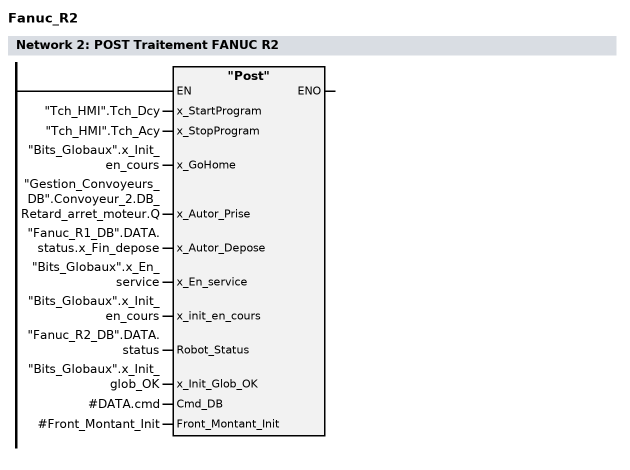
   RUNG wire#powerrail
      "Post"(x_StartProgram := "Tch_HMI".Tch_Dcy, x_StopProgram := "Tch_HMI".Tch_Acy, x_GoHome := "Bits_Globaux".x_Init_en_cours, x_Autor_Prise := "Gestion_Convoyeurs_DB".Convoyeur_2.DB_Retard_arret_moteur.Q, x_Autor_Depose := "Fanuc_R1_DB".DATA.status.x_Fin_depose, x_En_service := "Bits_Globaux".x_En_service, x_init_en_cours := "Bits_Globaux".x_Init_en_cours, Robot_Status := "Fanuc_R2_DB".DATA.status, x_Init_Glob_OK := "Bits_Globaux".x_Init_glob_OK, Cmd_DB := #DATA.cmd, Front_Montant_Init := #Front_Montant_Init)
   END_RUNG
   // the same network as SCL:
   "Post"(x_StartProgram := "Tch_HMI".Tch_Dcy,
          x_StopProgram := "Tch_HMI".Tch_Acy,
          x_GoHome := "Bits_Globaux".x_Init_en_cours,
          x_Autor_Prise := "Gestion_Convoyeurs_DB".Convoyeur_2.DB_Retard_arret_moteur.Q,
          x_Autor_Depose := "Fanuc_R1_DB".DATA.status.x_Fin_depose,
          x_En_service := "Bits_Globaux".x_En_service,
          x_init_en_cours := "Bits_Globaux".x_Init_en_cours,
          Robot_Status := "Fanuc_R2_DB".DATA.status,
          x_Init_Glob_OK := "Bits_Globaux".x_Init_glob_OK,
          Cmd_DB := #DATA.cmd,
          Front_Montant_Init := #Front_Montant_Init);
END_REGION
END_FUNCTION_BLOCK

// folder: 5-Cellule_conditionnement/GoFa_ABB_R3

FUNCTION_BLOCK "GoFa_R3_FB"   // FB15, LAD
TITLE = Commande ABB
{ S7_Optimized_Access := 'TRUE' }
VERSION : 0.1
   VAR
      GoFa_Status : "GoFa_Status";
      GoFa_Cmd : "GoFa_cmd";
      x_Demande_ecriture_Modbus : Bool;
   END_VAR
BEGIN

REGION Network 1: Allumage des moteurs
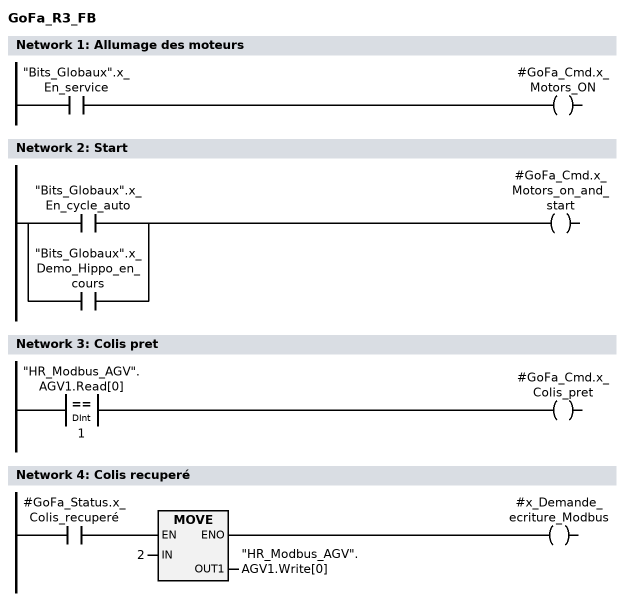
   RUNG wire#powerrail
      Contact( "Bits_Globaux".x_En_service )
      Coil( #GoFa_Cmd.x_Motors_ON )
   END_RUNG
   // the same network as SCL:
   #GoFa_Cmd.x_Motors_ON := "Bits_Globaux".x_En_service;
END_REGION

REGION Network 2: Start
   RUNG wire#powerrail
      Contact( "Bits_Globaux".x_En_cycle_auto )
      wire#w1
      Coil( #GoFa_Cmd.x_Motors_on_and_start )
   END_RUNG
   RUNG wire#powerrail
      Contact( "Bits_Globaux".x_Demo_Hippo_en_cours )
   END_RUNG wire#w1
   // the same network as SCL:
   #GoFa_Cmd.x_Motors_on_and_start := "Bits_Globaux".x_En_cycle_auto OR "Bits_Globaux".x_Demo_Hippo_en_cours;
END_REGION

REGION Network 3: Colis pret
   RUNG wire#powerrail
      { S7_Templates := "SrcType := DInt" } EQ_Contact(in1 := "HR_Modbus_AGV".AGV1.Read[0], in2 := 1)
      Coil( #GoFa_Cmd.x_Colis_pret )
   END_RUNG
   // the same network as SCL:
   #GoFa_Cmd.x_Colis_pret := "HR_Modbus_AGV".AGV1.Read[0] = 1;
END_REGION

REGION Network 4: Colis recuperé
   RUNG wire#powerrail
      Contact( #GoFa_Status.x_Colis_recuperé )
      Move(in := 2, out1 => "HR_Modbus_AGV".AGV1.Write[0])
      Coil( #x_Demande_ecriture_Modbus )
   END_RUNG
   // the same network as SCL:
   IF #GoFa_Status.x_Colis_recuperé THEN "HR_Modbus_AGV".AGV1.Write[0] := 2; END_IF;
   #x_Demande_ecriture_Modbus := #GoFa_Status.x_Colis_recuperé;
END_REGION
END_FUNCTION_BLOCK

// folder: 6_UR10_R5

FUNCTION_BLOCK "60_UR_R5"   // FB6, LAD
{ S7_Optimized_Access := 'TRUE' }
VERSION : 0.1
   VAR
      DATA : "UR_Cobot";
      x_DemandeEcriture_Modbus_AGV : Bool;
   END_VAR
   // // DATA.Registers_Out_2.Bits.Register[0] : Demande Init
   // // DATA.Registers_Out_2.Bits.Register[1] : EnCycleAuto
   // // DATA.Registers_Out_2.Bits.Register[2] : EnCycleDemo
   // // DATA.Registers_Out_2.Bits.Register[3] : PauseProgPLC
   // // DATA.Registers_Out_2.Bits.Register[4] : StopProgPLC
   // // DATA.Registers_Out_2.Bits.Register[5] : StartProgPLC (demarrage boucle Main)
   // // DATA.Registers_Out_2.Bits.Register[6] : Initialisation auto après AU
   // // DATA.Registers_Out_2.Bits.Register[7] : InitRequired
   // // DATA.Registers_Out_1.Bits.Register[0] : BoitePleineDispo
   // // DATA.Registers_Out_1.Bits.Register[1] : CouvercleDispo
   // // DATA.Registers_Out_1.Bits.Register[2] : AGVenPosition
   // // DATA.Registers.Bit.Register[0] : IsInitialized
   // // DATA.Registers.Bit.Register[1] : PriseOK
   // // DATA.Registers.Bit.Register[2] : DeposeOK
   // // DATA.Registers_Out_2.Bits.Register[8] : UnpauseProgPLC
BEGIN

REGION Network 1: Init Required?
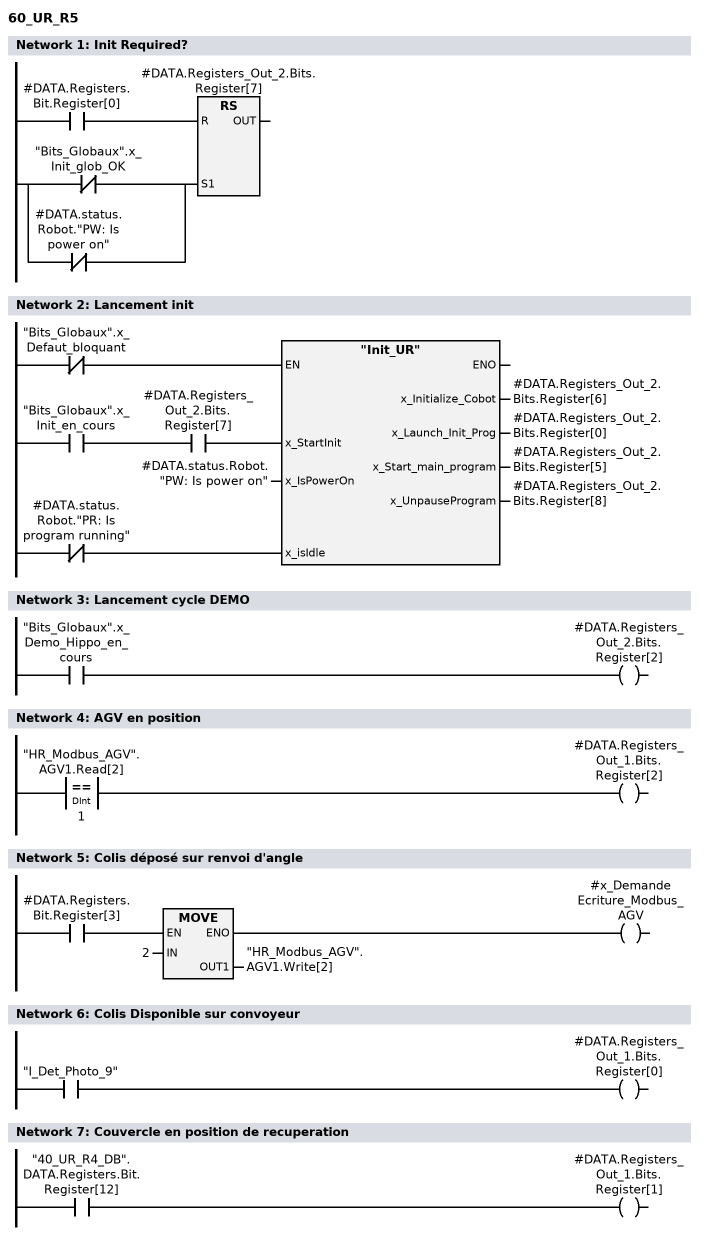
   RUNG wire#powerrail
      Contact( #DATA.Registers.Bit.Register[0] )
      S_RS(operand := #DATA.Registers_Out_2.Bits.Register[7], s1 := wire#w1)
   END_RUNG
   RUNG wire#powerrail
      I_Contact( "Bits_Globaux".x_Init_glob_OK )
   END_RUNG wire#w1
   RUNG wire#powerrail
      I_Contact( #DATA.status.Robot."PW: Is power on" )
   END_RUNG wire#w1
   // the same network as SCL:
   IF #DATA.Registers.Bit.Register[0] THEN
       #DATA.Registers_Out_2.Bits.Register[7] := FALSE;   // RS flip-flop
   END_IF;
   IF NOT "Bits_Globaux".x_Init_glob_OK OR NOT #DATA.status.Robot."PW: Is power on" THEN
       #DATA.Registers_Out_2.Bits.Register[7] := TRUE;
   END_IF;
END_REGION

REGION Network 2: Lancement init
   RUNG wire#powerrail
      I_Contact( "Bits_Globaux".x_Defaut_bloquant )
      "Init_UR"(x_StartInit := wire#w1, x_isIdle := wire#w2, x_IsPowerOn := #DATA.status.Robot."PW: Is power on", x_Initialize_Cobot => #DATA.Registers_Out_2.Bits.Register[6], x_Launch_Init_Prog => #DATA.Registers_Out_2.Bits.Register[0], x_Start_main_program => #DATA.Registers_Out_2.Bits.Register[5], x_UnpauseProgram => #DATA.Registers_Out_2.Bits.Register[8])
   END_RUNG
   RUNG wire#powerrail
      Contact( "Bits_Globaux".x_Init_en_cours )
      Contact( #DATA.Registers_Out_2.Bits.Register[7] )
   END_RUNG wire#w1
   RUNG wire#powerrail
      I_Contact( #DATA.status.Robot."PR: Is program running" )
   END_RUNG wire#w2
   // the same network as SCL:
   IF NOT "Bits_Globaux".x_Defaut_bloquant THEN
       "Init_UR"(x_StartInit := "Bits_Globaux".x_Init_en_cours AND #DATA.Registers_Out_2.Bits.Register[7],
                 x_IsPowerOn := #DATA.status.Robot."PW: Is power on",
                 x_isIdle := NOT #DATA.status.Robot."PR: Is program running",
                 x_Initialize_Cobot => #DATA.Registers_Out_2.Bits.Register[6],
                 x_Launch_Init_Prog => #DATA.Registers_Out_2.Bits.Register[0],
                 x_Start_main_program => #DATA.Registers_Out_2.Bits.Register[5],
                 x_UnpauseProgram => #DATA.Registers_Out_2.Bits.Register[8]);
   END_IF;
END_REGION

REGION Network 3: Lancement cycle DEMO
   RUNG wire#powerrail
      Contact( "Bits_Globaux".x_Demo_Hippo_en_cours )
      Coil( #DATA.Registers_Out_2.Bits.Register[2] )
   END_RUNG
   // the same network as SCL:
   #DATA.Registers_Out_2.Bits.Register[2] := "Bits_Globaux".x_Demo_Hippo_en_cours;
END_REGION

REGION Network 4: AGV en position
   RUNG wire#powerrail
      { S7_Templates := "SrcType := DInt" } EQ_Contact(in1 := "HR_Modbus_AGV".AGV1.Read[2], in2 := 1)
      Coil( #DATA.Registers_Out_1.Bits.Register[2] )
   END_RUNG
   // the same network as SCL:
   #DATA.Registers_Out_1.Bits.Register[2] := "HR_Modbus_AGV".AGV1.Read[2] = 1;
END_REGION

REGION Network 5: Colis déposé sur renvoi d'angle
   RUNG wire#powerrail
      Contact( #DATA.Registers.Bit.Register[3] )
      Move(in := 2, out1 => "HR_Modbus_AGV".AGV1.Write[2])
      Coil( #x_DemandeEcriture_Modbus_AGV )
   END_RUNG
   // the same network as SCL:
   IF #DATA.Registers.Bit.Register[3] THEN "HR_Modbus_AGV".AGV1.Write[2] := 2; END_IF;
   #x_DemandeEcriture_Modbus_AGV := #DATA.Registers.Bit.Register[3];
END_REGION

REGION Network 6: Colis Disponible sur convoyeur
   RUNG wire#powerrail
      Contact( "I_Det_Photo_9" )
      Coil( #DATA.Registers_Out_1.Bits.Register[0] )
   END_RUNG
   // the same network as SCL:
   #DATA.Registers_Out_1.Bits.Register[0] := "I_Det_Photo_9";
END_REGION

REGION Network 7: Couvercle en position de recuperation
   RUNG wire#powerrail
      Contact( "40_UR_R4_DB".DATA.Registers.Bit.Register[12] )
      Coil( #DATA.Registers_Out_1.Bits.Register[1] )
   END_RUNG
   // the same network as SCL:
   #DATA.Registers_Out_1.Bits.Register[1] := "40_UR_R4_DB".DATA.Registers.Bit.Register[12];
END_REGION
END_FUNCTION_BLOCK

// folder: 7_AGVs

FUNCTION_BLOCK "AGV_1"   // FB16, LAD
{ S7_Optimized_Access := 'TRUE' }
VERSION : 0.1
BEGIN

REGION Network 1: Com lancement Boucle grand colis vers ABB
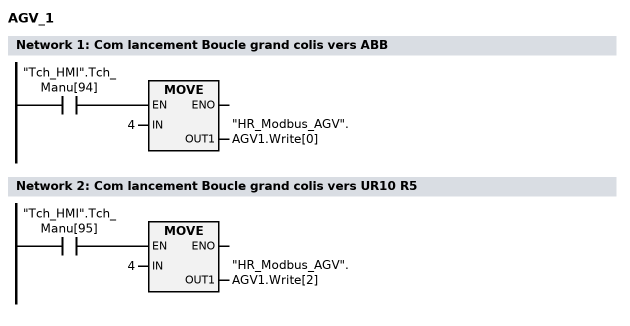
   RUNG wire#powerrail
      Contact( "Tch_HMI".Tch_Manu[94] )
      Move(in := 4, out1 => "HR_Modbus_AGV".AGV1.Write[0])
   END_RUNG
   // the same network as SCL:
   IF "Tch_HMI".Tch_Manu[94] THEN "HR_Modbus_AGV".AGV1.Write[0] := 4; END_IF;
END_REGION

REGION Network 2: Com lancement Boucle grand colis vers UR10 R5
   RUNG wire#powerrail
      Contact( "Tch_HMI".Tch_Manu[95] )
      Move(in := 4, out1 => "HR_Modbus_AGV".AGV1.Write[2])
   END_RUNG
   // the same network as SCL:
   IF "Tch_HMI".Tch_Manu[95] THEN "HR_Modbus_AGV".AGV1.Write[2] := 4; END_IF;
END_REGION
END_FUNCTION_BLOCK

FUNCTION_BLOCK "AGV_2"   // FB17, LAD
{ S7_Optimized_Access := 'TRUE' }
VERSION : 0.1
BEGIN

REGION Network 1: COM Lancement Boucle PC AGV2
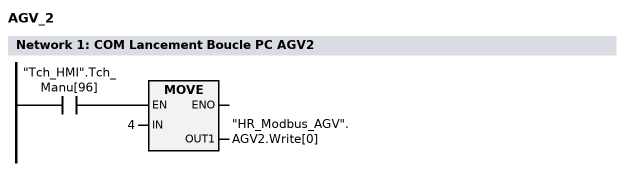
   RUNG wire#powerrail
      Contact( "Tch_HMI".Tch_Manu[96] )
      Move(in := 4, out1 => "HR_Modbus_AGV".AGV2.Write[0])
   END_RUNG
   // the same network as SCL:
   IF "Tch_HMI".Tch_Manu[96] THEN "HR_Modbus_AGV".AGV2.Write[0] := 4; END_IF;
END_REGION
END_FUNCTION_BLOCK

FUNCTION_BLOCK "AGVs_Modbus_Read_COM"   // FB18, LAD
{ S7_Optimized_Access := 'TRUE' }
VERSION : 0.1
   VAR
      MB_CLIENT_AGV1 : MB_CLIENT;
      MB_CLIENT_AGV2 : MB_CLIENT;
   END_VAR
BEGIN

REGION Network 1: Client modbus AGV1 read
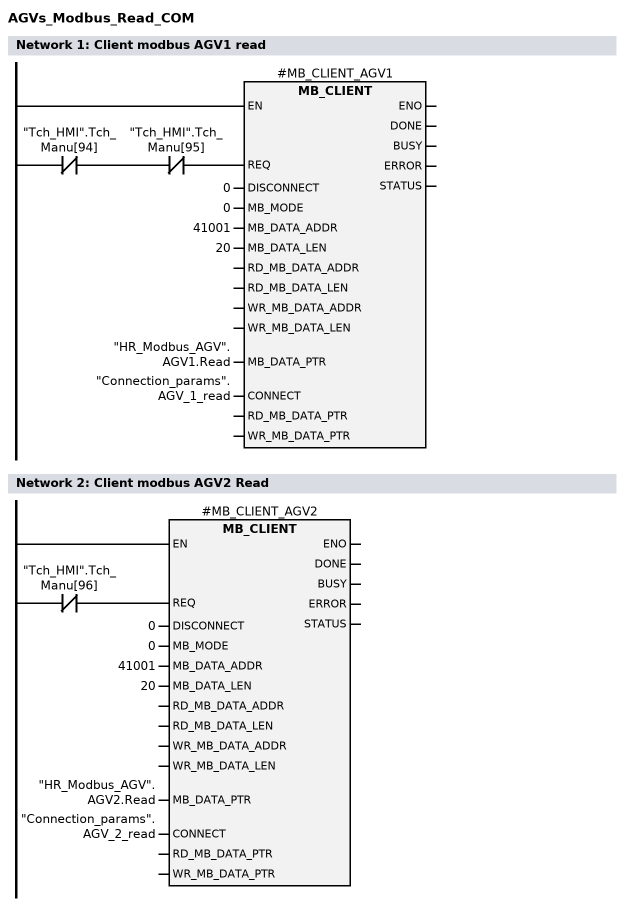
   #MB_CLIENT_AGV1(REQ := NOT "Tch_HMI".Tch_Manu[94] AND NOT "Tch_HMI".Tch_Manu[95],   // MB_CLIENT
                   DISCONNECT := 0,
                   MB_MODE := 0,
                   MB_DATA_ADDR := 41001,
                   MB_DATA_LEN := 20,
                   MB_DATA_PTR := "HR_Modbus_AGV".AGV1.Read,
                   CONNECT := "Connection_params".AGV_1_read);
END_REGION

REGION Network 2: Client modbus AGV2 Read
   #MB_CLIENT_AGV2(REQ := NOT "Tch_HMI".Tch_Manu[96],   // MB_CLIENT
                   DISCONNECT := 0,
                   MB_MODE := 0,
                   MB_DATA_ADDR := 41001,
                   MB_DATA_LEN := 20,
                   MB_DATA_PTR := "HR_Modbus_AGV".AGV2.Read,
                   CONNECT := "Connection_params".AGV_2_read);
END_REGION
END_FUNCTION_BLOCK

FUNCTION_BLOCK "AGVs_Modbus_Write_COM"   // FB19, LAD
{ S7_Optimized_Access := 'TRUE' }
VERSION : 0.1
   VAR
      MB_CLIENT_AGV1 : MB_CLIENT;
      MB_CLIENT_AGV2 : MB_CLIENT;
      DmdEcritureAGV1 : Bool;
      DmdEcritureAGV2 : Bool;
   END_VAR
BEGIN

REGION Network 1: INIT
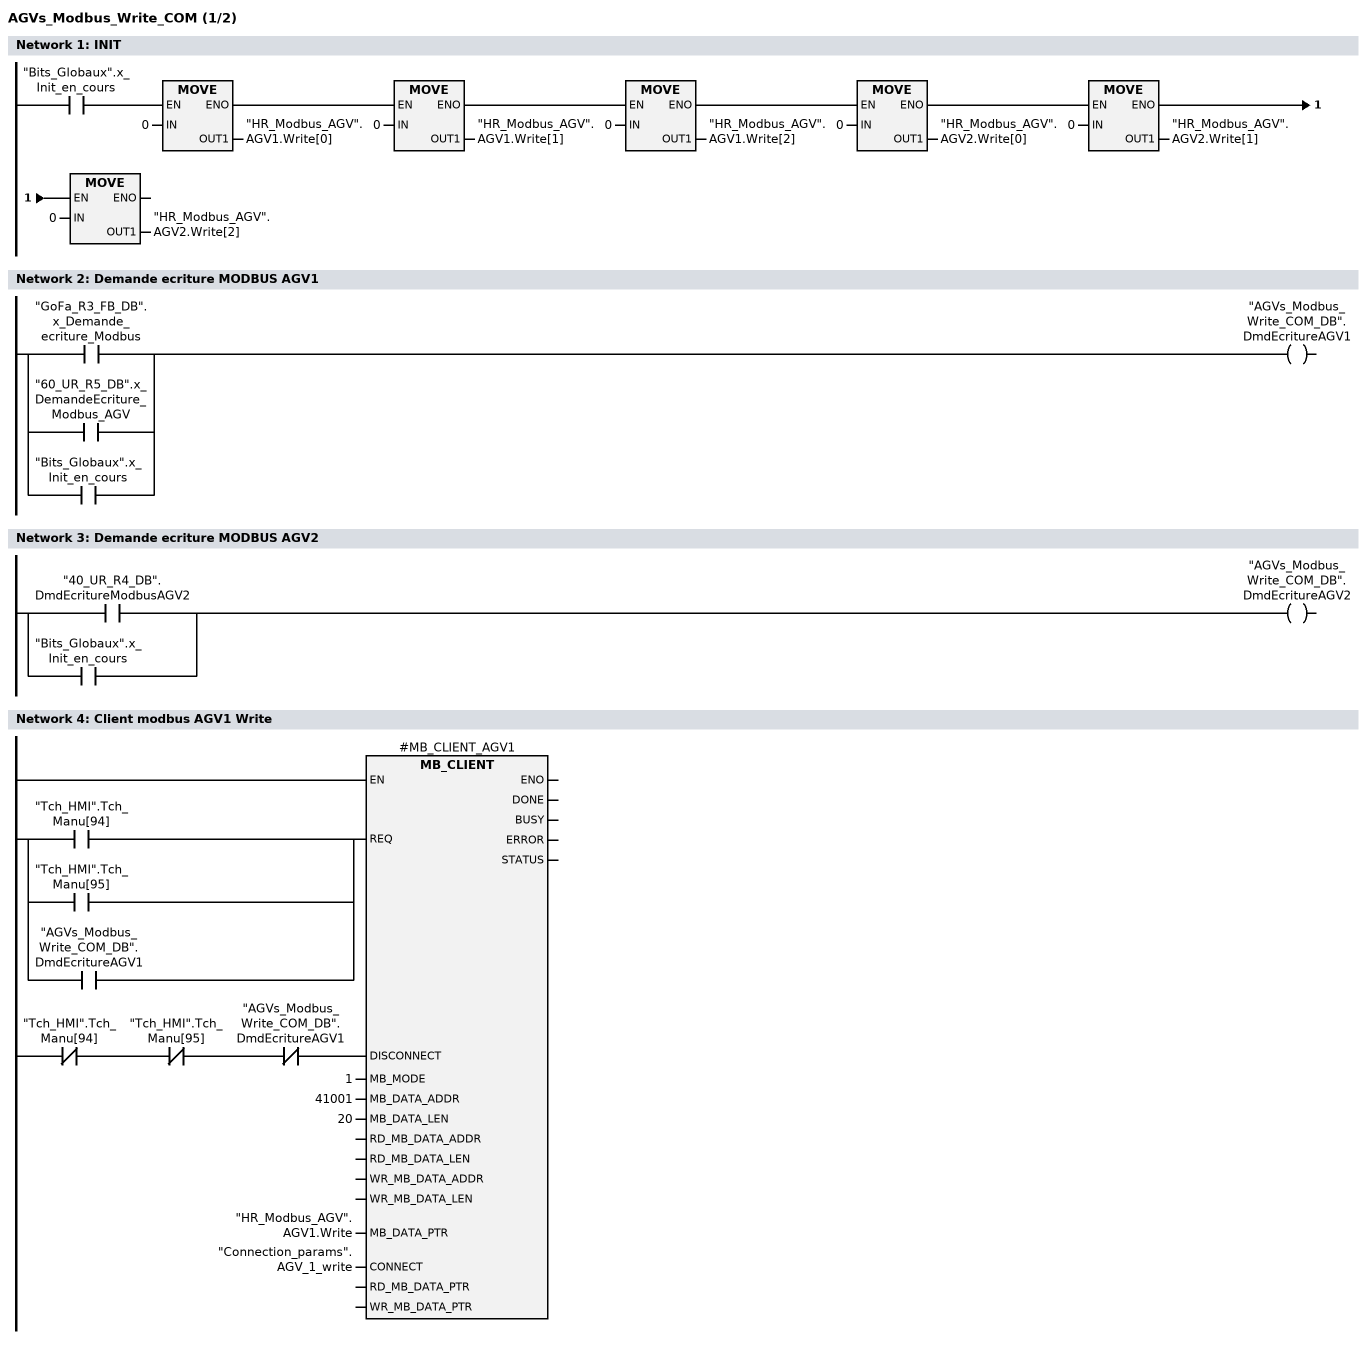
   RUNG wire#powerrail
      Contact( "Bits_Globaux".x_Init_en_cours )
      Move(in := 0, out1 => "HR_Modbus_AGV".AGV1.Write[0])
      Move(in := 0, out1 => "HR_Modbus_AGV".AGV1.Write[1])
      Move(in := 0, out1 => "HR_Modbus_AGV".AGV1.Write[2])
      Move(in := 0, out1 => "HR_Modbus_AGV".AGV2.Write[0])
      Move(in := 0, out1 => "HR_Modbus_AGV".AGV2.Write[1])
      Move(in := 0, out1 => "HR_Modbus_AGV".AGV2.Write[2])
   END_RUNG
   // the same network as SCL:
   IF "Bits_Globaux".x_Init_en_cours THEN
       "HR_Modbus_AGV".AGV1.Write[0] := 0;
       "HR_Modbus_AGV".AGV1.Write[1] := 0;
       "HR_Modbus_AGV".AGV1.Write[2] := 0;
       "HR_Modbus_AGV".AGV2.Write[0] := 0;
       "HR_Modbus_AGV".AGV2.Write[1] := 0;
       "HR_Modbus_AGV".AGV2.Write[2] := 0;
   END_IF;
END_REGION

REGION Network 2: Demande ecriture MODBUS AGV1
   RUNG wire#powerrail
      Contact( "GoFa_R3_FB_DB".x_Demande_ecriture_Modbus )
      wire#w1
      Coil( "AGVs_Modbus_Write_COM_DB".DmdEcritureAGV1 )
   END_RUNG
   RUNG wire#powerrail
      Contact( "60_UR_R5_DB".x_DemandeEcriture_Modbus_AGV )
   END_RUNG wire#w1
   RUNG wire#powerrail
      Contact( "Bits_Globaux".x_Init_en_cours )
   END_RUNG wire#w1
   // the same network as SCL:
   "AGVs_Modbus_Write_COM_DB".DmdEcritureAGV1 := "GoFa_R3_FB_DB".x_Demande_ecriture_Modbus OR "60_UR_R5_DB".x_DemandeEcriture_Modbus_AGV OR "Bits_Globaux".x_Init_en_cours;
END_REGION

REGION Network 3: Demande ecriture MODBUS AGV2
   RUNG wire#powerrail
      Contact( "40_UR_R4_DB".DmdEcritureModbusAGV2 )
      wire#w1
      Coil( "AGVs_Modbus_Write_COM_DB".DmdEcritureAGV2 )
   END_RUNG
   RUNG wire#powerrail
      Contact( "Bits_Globaux".x_Init_en_cours )
   END_RUNG wire#w1
   // the same network as SCL:
   "AGVs_Modbus_Write_COM_DB".DmdEcritureAGV2 := "40_UR_R4_DB".DmdEcritureModbusAGV2 OR "Bits_Globaux".x_Init_en_cours;
END_REGION

REGION Network 4: Client modbus AGV1 Write
   #MB_CLIENT_AGV1(REQ := "Tch_HMI".Tch_Manu[94] OR "Tch_HMI".Tch_Manu[95] OR "AGVs_Modbus_Write_COM_DB".DmdEcritureAGV1,   // MB_CLIENT
                   DISCONNECT := NOT "Tch_HMI".Tch_Manu[94] AND NOT "Tch_HMI".Tch_Manu[95] AND NOT "AGVs_Modbus_Write_COM_DB".DmdEcritureAGV1,
                   MB_MODE := 1,
                   MB_DATA_ADDR := 41001,
                   MB_DATA_LEN := 20,
                   MB_DATA_PTR := "HR_Modbus_AGV".AGV1.Write,
                   CONNECT := "Connection_params".AGV_1_write);
END_REGION

REGION Network 5: Client modbus AGV2 Write
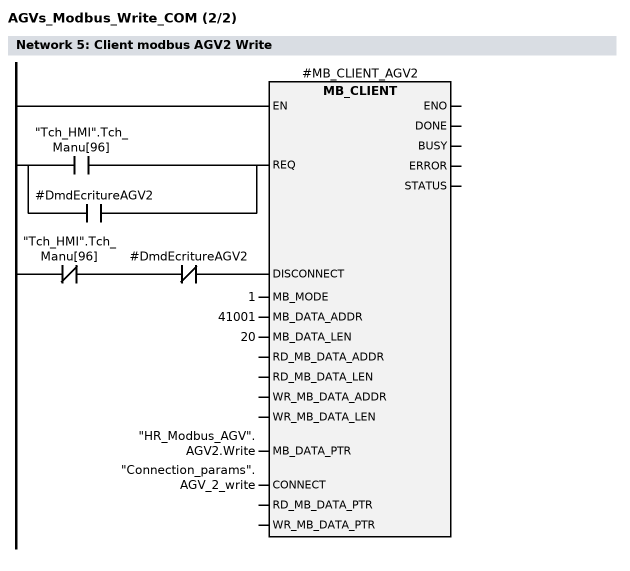
   #MB_CLIENT_AGV2(REQ := "Tch_HMI".Tch_Manu[96] OR #DmdEcritureAGV2,   // MB_CLIENT
                   DISCONNECT := NOT "Tch_HMI".Tch_Manu[96] AND NOT #DmdEcritureAGV2,
                   MB_MODE := 1,
                   MB_DATA_ADDR := 41001,
                   MB_DATA_LEN := 20,
                   MB_DATA_PTR := "HR_Modbus_AGV".AGV2.Write,
                   CONNECT := "Connection_params".AGV_2_write);
END_REGION
END_FUNCTION_BLOCK

// folder: 8_Alarmes

FUNCTION_BLOCK "Defauts"   // FB20, LAD
{ S7_Optimized_Access := 'TRUE' }
VERSION : 0.1
   VAR
      DB_Alarmes_hippodrome : "Create_Alarm";
      "Erreur elevateur hippodrome" : Array[0..1] of String;
   END_VAR
BEGIN

REGION Network 1: Defauts hippodrome
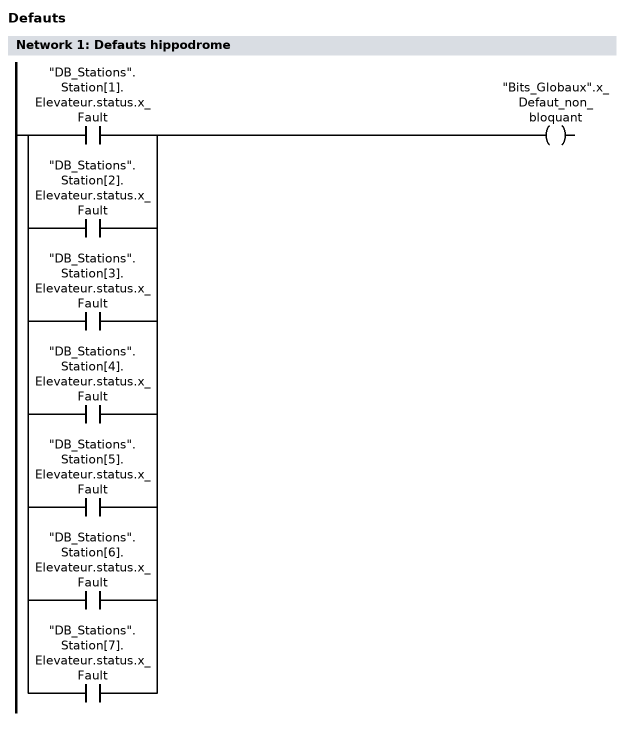
   RUNG wire#powerrail
      Contact( "DB_Stations".Station[1].Elevateur.status.x_Fault )
      wire#w1
      Coil( "Bits_Globaux".x_Defaut_non_bloquant )
   END_RUNG
   RUNG wire#powerrail
      Contact( "DB_Stations".Station[2].Elevateur.status.x_Fault )
   END_RUNG wire#w1
   RUNG wire#powerrail
      Contact( "DB_Stations".Station[3].Elevateur.status.x_Fault )
   END_RUNG wire#w1
   RUNG wire#powerrail
      Contact( "DB_Stations".Station[4].Elevateur.status.x_Fault )
   END_RUNG wire#w1
   RUNG wire#powerrail
      Contact( "DB_Stations".Station[5].Elevateur.status.x_Fault )
   END_RUNG wire#w1
   RUNG wire#powerrail
      Contact( "DB_Stations".Station[6].Elevateur.status.x_Fault )
   END_RUNG wire#w1
   RUNG wire#powerrail
      Contact( "DB_Stations".Station[7].Elevateur.status.x_Fault )
   END_RUNG wire#w1
   // the same network as SCL:
   "Bits_Globaux".x_Defaut_non_bloquant := "DB_Stations".Station[1].Elevateur.status.x_Fault OR "DB_Stations".Station[2].Elevateur.status.x_Fault OR "DB_Stations".Station[3].Elevateur.status.x_Fault OR "DB_Stations".Station[4].Elevateur.status.x_Fault OR "DB_Stations".Station[5].Elevateur.status.x_Fault OR "DB_Stations".Station[6].Elevateur.status.x_Fault OR "DB_Stations".Station[7].Elevateur.status.x_Fault;
END_REGION

REGION Network 2: Defauts canal 03
END_REGION
END_FUNCTION_BLOCK

(* ===== HMI "HMI_RT_1" =====
system functions are stored by id; their names below are inferred from use
connection "HMI_Liaison_1": ETHERNET, S7_1500_OMS

HMI tags "Table de variables standard"
   "Touche_Tch_FDCY" : Bool = PLC Tch_HMI.Tch_Acy, 1 s
   "Bits_B_Acy" : Bool = PLC Tch_HMI.Tch_Acy, 1 s
   "Bits_B_Dcy" : Bool = PLC Tch_HMI.Tch_Dcy, 1 s
   "I_En_Arret_Urgence" : Bool = PLC I_Not_AU AT %I0.1, 1 s
   "I_En_Automatique" : Bool = PLC I_En_Automatique AT %I0.3, 1 s
   "I_En_Service" : Bool = PLC I_En_Service AT %I0.0, 1 s
   "Touche_Tch_DCY" : Bool = PLC Tch_HMI.Tch_Dcy, 1 s
   "Bits_B_defaut_en_cours" : Bool = PLC Bits_Globaux.x_Defaut_bloquant, 1 s
   "I_En_Manuel" : Bool = PLC I_En_Manuel AT %I0.2, 1 s
   "I_porte_non_réarmée" : Bool = PLC I_porte_non_réarmée AT %I0.4, 1 s
   "I_porte_01_Op" : Bool = PLC I_porte_01_Op AT %I0.5, 1 s
   "I_porte_02_Op" : Bool = PLC I_porte_02_Op AT %I0.6, 1 s
   "I_libre_I07" : Bool = PLC I_libre_I07 AT %I0.7, 1 s
   "I_libre_I10" : Bool = PLC I_libre_I10 AT %I1.0, 1 s
   "I_Def_Thermique_CV01_hyppo" : Bool = PLC I_Def_Thermique_CV01_hyppo AT %I1.1, 1 s
   "I_Def_Thermique_CV02_hyppo" : Bool = PLC I_Def_Thermique_CV02_hyppo AT %I1.2, 1 s
   "I_Def_Thermique_CV03_hyppo" : Bool = PLC I_Def_Thermique_CV03_hyppo AT %I1.3, 1 s
   "I_Def_Thermique_CV04_hyppo" : Bool = PLC I_Def_Thermique_CV04_hyppo AT %I1.4, 1 s
   "I_libre_I15" : Bool = PLC I_libre_I15 AT %I1.5, 1 s
   "I_libre_I16" : Bool = PLC I_libre_I16 AT %I1.6, 1 s
   "I_libre_I17" : Bool = PLC I_libre_I17 AT %I1.7, 1 s
   "I_libre_I20" : Bool = PLC I_libre_I20 AT %I2.0, 1 s
   "I_libre_I21" : Bool = PLC I_libre_I21 AT %I2.1, 1 s
   "I_libre_I22" : Bool = PLC I_libre_I22 AT %I2.2, 1 s
   "I_libre_I23" : Bool = PLC I_libre_I23 AT %I2.3, 1 s
   "I_libre_I24" : Bool = PLC I_libre_I24 AT %I2.4, 1 s
   "I_libre_I25" : Bool = PLC I_libre_I25 AT %I2.5, 1 s
   "I_libre_I26" : Bool = PLC I_libre_I26 AT %I2.6, 1 s
   "I_libre_I27" : Bool = PLC I_libre_I27 AT %I2.7, 1 s
   "I_libre_I30" : Bool = PLC I_libre_I30 AT %I3.0, 1 s
   "I_libre_I31" : Bool = PLC I_libre_I31 AT %I3.1, 1 s
   "I_libre_I32" : Bool = PLC I_libre_I32 AT %I3.2, 1 s
   "I_libre_I33" : Bool = PLC I_libre_I33 AT %I3.3, 1 s
   "I_libre_I34" : Bool = PLC I_libre_I34 AT %I3.4, 1 s
   "I_libre_I35" : Bool = PLC I_libre_I35 AT %I3.5, 1 s
   "I_libre_I36" : Bool = PLC I_libre_I36 AT %I3.6, 1 s
   "I_libre_I37" : Bool = PLC I_libre_I37 AT %I3.7, 1 s
   "Q_CL_verte" : Bool = PLC O_CL_verte AT %Q0.0, 1 s
   "Q_CL_Orange" : Bool = PLC O_CL_Orange AT %Q0.1, 1 s
   "Q_CL_Rouge" : Bool = PLC O_CL_Rouge AT %Q0.2, 1 s
   "Q_LibreQ03" : Bool = PLC Q_LibreQ03 AT %Q0.3, 1 s
   "Q_LibreQ04" : Bool = PLC Q_LibreQ04 AT %Q0.4, 1 s
   "Q_LibreQ05" : Bool = PLC Q_LibreQ05 AT %Q0.5, 1 s
   "Q_LibreQ06" : Bool = PLC Q_LibreQ06 AT %Q0.6, 1 s
   "Q_LibreQ07" : Bool = PLC Q_LibreQ07 AT %Q0.7, 1 s
   "Q_LibreQ10" : Bool = PLC Q_LibreQ10 AT %Q1.0, 1 s
   "Q_LibreQ11" : Bool = PLC Q_LibreQ11 AT %Q1.1, 1 s
   "Q_LibreQ12" : Bool = PLC Q_LibreQ12 AT %Q1.2, 1 s
   "Q_LibreQ13" : Bool = PLC Q_LibreQ13 AT %Q1.3, 1 s
   "Q_LibreQ14" : Bool = PLC Q_LibreQ14 AT %Q1.4, 1 s
   "Q_LibreQ15" : Bool = PLC Q_LibreQ15 AT %Q1.5, 1 s
   "Q_LibreQ16" : Bool = PLC Q_LibreQ16 AT %Q1.6, 1 s
   "Q_LibreQ17" : Bool = PLC Q_LibreQ17 AT %Q1.7, 1 s
   "Q_LibreQ24" : Bool = PLC Q_LibreQ24 AT %Q2.4, 1 s
   "Q_LibreQ25" : Bool = PLC Q_LibreQ25 AT %Q2.5, 1 s
   "Q_LibreQ26" : Bool = PLC Q_LibreQ26 AT %Q2.6, 1 s
   "Q_LibreQ27" : Bool = PLC Q_LibreQ27 AT %Q2.7, 1 s
   "Q_LibreQ30" : Bool = PLC Q_LibreQ30 AT %Q3.0, 1 s
   "Q_LibreQ31" : Bool = PLC Q_LibreQ31 AT %Q3.1, 1 s
   "Q_LibreQ32" : Bool = PLC Q_LibreQ32 AT %Q3.2, 1 s
   "Q_LibreQ33" : Bool = PLC Q_LibreQ33 AT %Q3.3, 1 s
   "Q_LibreQ34" : Bool = PLC Q_LibreQ34 AT %Q3.4, 1 s
   "Q_LibreQ35" : Bool = PLC Q_LibreQ35 AT %Q3.5, 1 s
   "Q_LibreQ37" : Bool = PLC Q_LibreQ37 AT %Q3.7, 1 s
   "Q_LibreQ36" : Bool = PLC Q_LibreQ36 AT %Q3.6, 1 s
   "Q_ON_CV_01_Hyppo" : Bool = PLC O_ON_CV_01_Hyppo AT %Q2.0, 1 s
   "Q_ON_CV_02_Hyppo" : Bool = PLC O_ON_CV_02_Hyppo AT %Q2.1, 1 s
   "Q_ON_CV_03_Hyppo" : Bool = PLC O_ON_CV_03_Hyppo AT %Q2.2, 1 s
   "Q_ON_CV_04_Hyppo" : Bool = PLC O_ON_CV_04_Hyppo AT %Q2.3, 1 s
   "I_Pres_Pal_B01" : Bool = PLC I_Pres_Pal_B01 AT %I5.0, 1 s
   "I_Pres_Elev_B01" : Bool = PLC I_Pres_Elev_B01 AT %I4.0, 1 s
   "I_Pres_Pal_B03" : Bool = PLC I_Pres_Pal_B03 AT %I5.4, 1 s
   "I_Elev_01_Bas" : Bool = PLC I_Elev_01_Bas AT %I5.1, 1 s
   "I_Elev_01_Haut" : Bool = PLC I_Elev_01_Haut AT %I4.1, 1 s
   "I_Pres_Pal_B02" : Bool = PLC I_Pres_Pal_B02 AT %I5.2, 1 s
   "I_Pres_Elev_B02" : Bool = PLC I_Pres_Elev_B02 AT %I4.2, 1 s
   "I_Elev_02_Bas" : Bool = PLC I_Elev_02_Bas AT %I5.3, 1 s
   "I_Elev_02_Haut" : Bool = PLC I_Elev_02_Haut AT %I4.3, 1 s
   "I_Pres_Pal_B04" : Bool = PLC I_Pres_Pal_B04 AT %I5.6, 1 s
   "I_Pres_Pal_B05" : Bool = PLC I_Pres_Pal_B05 AT %I7.0, 1 s
   "I_Pres_Pal_B06" : Bool = PLC I_Pres_Pal_B06 AT %I7.2, 1 s
   "I_Pres_Pal_B07" : Bool = PLC I_Pres_Pal_B07 AT %I7.4, 1 s
   "I_Pres_Elev_B03" : Bool = PLC I_Pres_Elev_B03 AT %I4.4, 1 s
   "I_Pres_Elev_B04" : Bool = PLC I_Pres_Elev_B04 AT %I4.6, 1 s
   "I_Pres_Elev_B05" : Bool = PLC I_Pres_Elev_B05 AT %I6.0, 1 s
   "I_Pres_Elev_B06" : Bool = PLC I_Pres_Elev_B06 AT %I6.2, 1 s
   "I_Pres_Elev_B07" : Bool = PLC I_Pres_Elev_B07 AT %I6.4, 1 s
   "I_Elev_03_Bas" : Bool = PLC I_Elev_03_Bas AT %I5.5, 1 s
   "I_Elev_03_Haut" : Bool = PLC I_Elev_03_Haut AT %I4.5, 1 s
   "I_Elev_04_Bas" : Bool = PLC I_Elev_04_Bas AT %I5.7, 1 s
   "I_Elev_04_Haut" : Bool = PLC I_Elev_04_Haut AT %I4.7, 1 s
   "I_Elev_05_Bas" : Bool = PLC I_Elev_05_Bas AT %I7.1, 1 s
   "I_Elev_05_Haut" : Bool = PLC I_Elev_05_Haut AT %I6.1, 1 s
   "I_Elev_06_Bas" : Bool = PLC I_Elev_06_Bas AT %I7.3, 1 s
   "I_Elev_06_Haut" : Bool = PLC I_Elev_06_Haut AT %I6.3, 1 s
   "I_Elev_07_Bas" : Bool = PLC I_Elev_07_Bas AT %I7.5, 1 s
   "I_Elev_07_Haut" : Bool = PLC I_Elev_07_Haut AT %I6.5, 1 s
   "AlwaysFALSE" : Bool = PLC AlwaysFALSE AT %M1.3, 1 s
   "Touche_Tch_Acquit" : Bool = PLC Tch_HMI.Tch_Acquit, 1 s
   "Touche_Tch_Manu{0}" : Bool = PLC Tch_HMI.Tch_Manu[0], 1 s
   "Touche_Tch_Manu{1}" : Bool = PLC Tch_HMI.Tch_Manu[1], 1 s
   "Touche_Tch_Manu{2}" : Bool = PLC Tch_HMI.Tch_Manu[2], 1 s
   "Touche_Tch_Manu{3}" : Bool = PLC Tch_HMI.Tch_Manu[3], 1 s
   "Touche_Tch_Manu{4}" : Bool = PLC Tch_HMI.Tch_Manu[4], 1 s
   "Touche_Tch_Manu{5}" : Bool = PLC Tch_HMI.Tch_Manu[5], 1 s
   "Touche_Tch_Manu{6}" : Bool = PLC Tch_HMI.Tch_Manu[6], 1 s
   "Touche_Tch_Manu{7}" : Bool = PLC Tch_HMI.Tch_Manu[7], 1 s
   "Touche_Tch_Manu{8}" : Bool = PLC Tch_HMI.Tch_Manu[8], 1 s
   "Touche_Tch_Manu{9}" : Bool = PLC Tch_HMI.Tch_Manu[9], 1 s
   "Touche_Tch_Manu{10}" : Bool = PLC Tch_HMI.Tch_Manu[10], 1 s
   "Touche_Tch_Manu{11}" : Bool = PLC Tch_HMI.Tch_Manu[11], 1 s
   "Touche_Tch_Manu{12}" : Bool = PLC Tch_HMI.Tch_Manu[12], 1 s
   "Touche_Tch_Manu{13}" : Bool = PLC Tch_HMI.Tch_Manu[13], 1 s
   "Touche_Tch_Manu{14}" : Bool = PLC Tch_HMI.Tch_Manu[14], 1 s
   "Touche_Tch_Manu{15}" : Bool = PLC Tch_HMI.Tch_Manu[15], 1 s
   "Touche_Tch_Manu{16}" : Bool = PLC Tch_HMI.Tch_Manu[16], 1 s
   "Touche_Tch_Manu{17}" : Bool = PLC Tch_HMI.Tch_Manu[17], 1 s
   "Touche_Tch_Manu{18}" : Bool = PLC Tch_HMI.Tch_Manu[18], 1 s
   "Touche_Tch_Manu{19}" : Bool = PLC Tch_HMI.Tch_Manu[19], 1 s
   "Touche_Tch_Manu{20}" : Bool = PLC Tch_HMI.Tch_Manu[20], 1 s
   "Touche_Tch_Manu{21}" : Bool = PLC Tch_HMI.Tch_Manu[21], 1 s
   "Touche_Tch_Manu{22}" : Bool = PLC Tch_HMI.Tch_Manu[22], 1 s
   "Touche_Tch_Manu{23}" : Bool = PLC Tch_HMI.Tch_Manu[23], 1 s
   "Touche_Tch_Manu{24}" : Bool = PLC Tch_HMI.Tch_Manu[24], 1 s
   "Touche_Tch_Manu{25}" : Bool = PLC Tch_HMI.Tch_Manu[25], 1 s
   "Touche_Tch_Manu{26}" : Bool = PLC Tch_HMI.Tch_Manu[26], 1 s
   "Touche_Tch_Manu{27}" : Bool = PLC Tch_HMI.Tch_Manu[27], 1 s
   "Touche_Tch_Manu{28}" : Bool = PLC Tch_HMI.Tch_Manu[28], 1 s
   "Touche_Tch_Manu{29}" : Bool = PLC Tch_HMI.Tch_Manu[29], 1 s
   "Touche_Tch_Manu{30}" : Bool = PLC Tch_HMI.Tch_Manu[30], 1 s
   "Touche_Tch_Manu{31}" : Bool = PLC Tch_HMI.Tch_Manu[31], 1 s
   "Touche_Tch_Manu{32}" : Bool = PLC Tch_HMI.Tch_Manu[32], 1 s
   "Touche_Tch_Manu{33}" : Bool = PLC Tch_HMI.Tch_Manu[33], 1 s
   "Touche_Tch_Manu{34}" : Bool = PLC Tch_HMI.Tch_Manu[34], 1 s
   "Touche_Tch_Manu{35}" : Bool = PLC Tch_HMI.Tch_Manu[35], 1 s
   "Touche_Tch_Manu{36}" : Bool = PLC Tch_HMI.Tch_Manu[36], 1 s
   "Touche_Tch_Manu{37}" : Bool = PLC Tch_HMI.Tch_Manu[37], 1 s
   "Touche_Tch_Manu{38}" : Bool = PLC Tch_HMI.Tch_Manu[38], 1 s
   "Touche_Tch_Manu{39}" : Bool = PLC Tch_HMI.Tch_Manu[39], 1 s
   "Touche_Tch_Manu{40}" : Bool = PLC Tch_HMI.Tch_Manu[40], 1 s
   "Touche_Tch_Manu{41}" : Bool = PLC Tch_HMI.Tch_Manu[41], 1 s
   "Touche_Tch_Manu{42}" : Bool = PLC Tch_HMI.Tch_Manu[42], 1 s
   "Touche_Tch_Manu{43}" : Bool = PLC Tch_HMI.Tch_Manu[43], 1 s
   "Touche_Tch_Manu{44}" : Bool = PLC Tch_HMI.Tch_Manu[44], 1 s
   "Touche_Tch_Manu{45}" : Bool = PLC Tch_HMI.Tch_Manu[45], 1 s
   "Touche_Tch_Manu{46}" : Bool = PLC Tch_HMI.Tch_Manu[46], 1 s
   "Touche_Tch_Manu{47}" : Bool = PLC Tch_HMI.Tch_Manu[47], 1 s
   "Touche_Tch_Manu{48}" : Bool = PLC Tch_HMI.Tch_Manu[48], 1 s
   "Touche_Tch_Manu{49}" : Bool = PLC Tch_HMI.Tch_Manu[49], 1 s
   "Touche_Tch_Manu{50}" : Bool = PLC Tch_HMI.Tch_Manu[50], 1 s
   "Touche_Tch_Manu{51}" : Bool = PLC Tch_HMI.Tch_Manu[51], 1 s
   "Touche_Tch_Manu{52}" : Bool = PLC Tch_HMI.Tch_Manu[52], 1 s
   "Touche_Tch_Manu{53}" : Bool = PLC Tch_HMI.Tch_Manu[53], 1 s
   "Touche_Tch_Manu{54}" : Bool = PLC Tch_HMI.Tch_Manu[54], 1 s
   "Touche_Tch_Manu{55}" : Bool = PLC Tch_HMI.Tch_Manu[55], 1 s
   "Touche_Tch_Manu{56}" : Bool = PLC Tch_HMI.Tch_Manu[56], 1 s
   "Touche_Tch_Manu{57}" : Bool = PLC Tch_HMI.Tch_Manu[57], 1 s
   "Touche_Tch_Manu{58}" : Bool = PLC Tch_HMI.Tch_Manu[58], 1 s
   "Touche_Tch_Manu{59}" : Bool = PLC Tch_HMI.Tch_Manu[59], 1 s
   "Touche_Tch_Manu{60}" : Bool = PLC Tch_HMI.Tch_Manu[60], 1 s
   "Touche_Tch_Manu{61}" : Bool = PLC Tch_HMI.Tch_Manu[61], 1 s
   "I_det_Phot_01" : Bool = PLC I_det_Phot_01 AT %I11.0, 1 s
   "I_det_Phot_02" : Bool = PLC I_det_Phot_02 AT %I10.0, 1 s
   "I_det_Phot_03" : Bool = PLC I_det_Phot_03 AT %I11.1, 1 s
   "I_verin_blocage_boite_rentré_01" : Bool = PLC I_verin_blocage_boite_rentré_01 AT %I11.2, 1 s
   "I_verin_blocage_boite_sorti_01" : Bool = PLC I_verin_blocage_boite_sorti_01 AT %I10.1, 1 s
   "I_verin_blocage_boite_sorti_02" : Bool = PLC I_verin_blocage_boite_sorti_02 AT %I10.2, 1 s
   "I_verin_blocage_boite_rentré_02" : Bool = PLC I_verin_blocage_boite_rentré_02 AT %I11.3, 1 s
   "I_verin_blocage_boite_sorti_03" : Bool = PLC I_verin_blocage_boite_sorti_03 AT %I10.3, 1 s
   "I_verin_blocage_boite_rentré_03" : Bool = PLC I_verin_blocage_boite_sorti_04 AT %I10.4, 1 s
   "I_verin_blocage_boite_sorti_04" : Bool = PLC I_verin_blocage_boite_rentré_03 AT %I11.4, 1 s
   "I_verin_blocage_boite_rentré_04" : Bool = PLC I_verin_blocage_boite_rentré_04 AT %I11.5, 1 s
   "I_det_photo_01" : Bool = PLC I_Det_Phot_04 AT %I13.0, 1 s
   "I_det_photo_02" : Bool = PLC I_Det_Phot_05 AT %I12.0, 1 s
   "I_det_photo_03" : Bool = PLC I_Det_Phot_06 AT %I13.1, 1 s
   "I_Det_Photo_7" : Bool = PLC I_Det_Photo_7 AT %I15.0, 1 s
   "I_Det_Photo_8" : Bool = PLC I_Det_Photo_8 AT %I14.0, 1 s
   "I_Det_Photo_9" : Bool = PLC I_Det_Photo_9 AT %I15.1, 1 s
   "Touche_Tch_Manu{62}" : Bool = PLC Tch_HMI.Tch_Manu[62], 1 s
   "Touche_Tch_Manu{63}" : Bool = PLC Tch_HMI.Tch_Manu[63], 1 s
   "Touche_Tch_Manu{64}" : Bool = PLC Tch_HMI.Tch_Manu[64], 1 s
   "Touche_Tch_Manu{65}" : Bool = PLC Tch_HMI.Tch_Manu[65], 1 s
   "Touche_Tch_Manu{66}" : Bool = PLC Tch_HMI.Tch_Manu[66], 1 s
   "Touche_Tch_Manu{67}" : Bool = PLC Tch_HMI.Tch_Manu[67], 1 s
   "O_Rentrer_Blocage_boite_01" : Bool = PLC O_Rentrer_Blocage_boite_01 AT %Q14.1, 1 s
   "O_Sortir_Blocage_boite_01" : Bool = PLC O_Sortir_Blocage_boite_01 AT %Q14.0, 1 s
   "O_Sortir_Blocage_boite_02" : Bool = PLC O_Sortir_Blocage_boite_02 AT %Q14.2, 1 s
   "O_Sortir_Blocage_boite_03" : Bool = PLC O_Sortir_Blocage_boite_03 AT %Q14.4, 1 s
   "O_Sortir_Blocage_boite_04" : Bool = PLC O_Sortir_Blocage_boite_04 AT %Q14.6, 1 s
   "O_Rentrer_Blocage_boite_02" : Bool = PLC O_Rentrer_Blocage_boite_02 AT %Q14.3, 1 s
   "O_Rentrer_Blocage_boite_03" : Bool = PLC O_Rentrer_Blocage_boite_03 AT %Q14.5, 1 s
   "O_Rentrer_Blocage_boite_04" : Bool = PLC O_Rentrer_Blocage_boite_04 AT %Q14.7, 1 s
   "O_Rentrer_Butée_01" : Bool = PLC O_Rentrer_Butée_01 AT %Q10.0, 1 s
   "O_Rentrer_Butée_02" : Bool = PLC O_Rentrer_Butée_02 AT %Q10.4, 1 s
   "O_Rentrer_Butée_03" : Bool = PLC O_Rentrer_Butée_03 AT %Q11.0, 1 s
   "O_Rentrer_Butée_04" : Bool = PLC O_Rentrer_Butée_04 AT %Q11.4, 1 s
   "O_Rentrer_Butée_05" : Bool = PLC O_Rentrer_Butée_05 AT %Q12.0, 1 s
   "O_Rentrer_Butée_06" : Bool = PLC O_Rentrer_Butée_06 AT %Q12.4, 1 s
   "O_Rentrer_Butée_07" : Bool = PLC O_Rentrer_Butée_07 AT %Q13.0, 1 s
   "O_Rentrer_Butée_EL_01" : Bool = PLC O_Rentrer_Butée_EL_01 AT %Q10.1, 1 s
   "O_Rentrer_Butée_EL_02" : Bool = PLC O_Rentrer_Butée_EL_02 AT %Q10.5, 1 s
   "O_Rentrer_Butée_EL_03" : Bool = PLC O_Rentrer_Butée_EL_03 AT %Q11.1, 1 s
   "O_Rentrer_Butée_EL_04" : Bool = PLC O_Rentrer_Butée_EL_04 AT %Q11.5, 1 s
   "O_Rentrer_Butée_EL_05" : Bool = PLC O_Rentrer_Butée_EL_05 AT %Q12.1, 1 s
   "O_Rentrer_Butée_EL_06" : Bool = PLC O_Rentrer_Butée_EL_06 AT %Q12.5, 1 s
   "O_Rentrer_Butée_EL_07" : Bool = PLC O_Rentrer_Butée_EL_07 AT %Q13.1, 1 s
   "O_Monter_EL_01" : Bool = PLC O_Monter_EL_01 AT %Q10.2, 1 s
   "O_Desc_EL_01" : Bool = PLC O_Desc_EL_01 AT %Q10.3, 1 s
   "O_Monter_EL_02" : Bool = PLC O_Monter_EL_02 AT %Q10.6, 1 s
   "O_Monter_EL_03" : Bool = PLC O_Monter_EL_03 AT %Q11.2, 1 s
   "O_Monter_EL_04" : Bool = PLC O_Monter_EL_04 AT %Q11.6, 1 s
   "O_Monter_EL_05" : Bool = PLC O_Monter_EL_05 AT %Q12.2, 1 s
   "O_Monter_EL_06" : Bool = PLC O_Monter_EL_06 AT %Q12.6, 1 s
   "O_Monter_EL_07" : Bool = PLC O_Monter_EL_07 AT %Q13.2, 1 s
   "O_Desc_EL_02" : Bool = PLC O_Desc_EL_02 AT %Q10.7, 1 s
   "O_Desc_EL_03" : Bool = PLC O_Desc_EL_03 AT %Q11.3, 1 s
   "O_Desc_EL_04" : Bool = PLC O_Desc_EL_04 AT %Q11.7, 1 s
   "O_Desc_EL_05" : Bool = PLC O_Desc_EL_05 AT %Q12.3, 1 s
   "O_Desc_EL_06" : Bool = PLC O_Desc_EL_06 AT %Q12.7, 1 s
   "O_Desc_EL_07" : Bool = PLC O_Desc_EL_07 AT %Q13.3, 1 s
   "O_Op_Porte_Vision" : Bool = PLC O_Op_Porte_Vision AT %Q13.4, 1 s
   "O_Cl_porte_Vision" : Bool = PLC O_Cl_porte_Vision AT %Q13.5, 1 s
   "Touche_Tch_Manu{68}" : Bool = PLC Tch_HMI.Tch_Manu[68], 1 s
   "Touche_Tch_Manu{69}" : Bool = PLC Tch_HMI.Tch_Manu[69], 1 s
   "Touche_Tch_Manu{70}" : Bool = PLC Tch_HMI.Tch_Manu[70], 1 s
   "Touche_Tch_Manu{71}" : Bool = PLC Tch_HMI.Tch_Manu[71], 1 s
   "Touche_Tch_Manu{80}" : Bool = PLC Tch_HMI.Tch_Manu[80], 1 s
   "Touche_Tch_Manu{81}" : Bool = PLC Tch_HMI.Tch_Manu[81], 1 s
   "Touche_Tch_Manu{82}" : Bool = PLC Tch_HMI.Tch_Manu[82], 1 s
   "Touche_Tch_Manu{83}" : Bool = PLC Tch_HMI.Tch_Manu[83], 1 s
   "Touche_Tch_Manu{84}" : Bool = PLC Tch_HMI.Tch_Manu[84], 1 s
   "Touche_Tch_Manu{85}" : Bool = PLC Tch_HMI.Tch_Manu[85], 1 s
   "Touche_Tch_Manu{86}" : Bool = PLC Tch_HMI.Tch_Manu[86], 1 s
   "Touche_Tch_Manu{87}" : Bool = PLC Tch_HMI.Tch_Manu[87], 1 s
   "Défauts_Def_Canal01" : Int = PLC Défauts.Def_Canal01 AT %DB13.DBW14, 1 s
   "Défauts_Def_Canal02" : Int = PLC Défauts.Def_Canal02 AT %DB13.DBW16, 1 s
   "Bits_B_Demo_Hyppo" : Bool = PLC Tch_HMI.Tch_Demo, 500 ms
   "Parametres_Sp_Vitesse_C01" : Int = PLC Parametres.Convoyeurs.Auto.i_Vitesse_C01, 1 s
   "Parametres_Sp_Vitesse_C02" : Int = PLC Parametres.Convoyeurs.Auto.i_Vitesse_C02, 1 s
   "Parametres_Sp_Vitesse_C03" : Int = PLC Parametres.Convoyeurs.Auto.i_Vitesse_C03, 1 s
   "Touche_Tch_Init" : Bool = PLC Tch_HMI.Tch_Init, 1 s
   "Défauts_Defauts{0}" : Bool = PLC Défauts.Defauts[0] AT %DB13.DBX0.0, 1 s
   "Défauts_Defauts{1}" : Bool = PLC Défauts.Defauts[1] AT %DB13.DBX0.1, 1 s
   "Défauts_Defauts{2}" : Bool = PLC Défauts.Defauts[2] AT %DB13.DBX0.2, 1 s
   "Défauts_Defauts{12}" : Bool = PLC Défauts.Defauts[12] AT %DB13.DBX1.4, 1 s
   "Défauts_Defauts{13}" : Bool = PLC Défauts.Defauts[13] AT %DB13.DBX1.5, 1 s
   "Défauts_Defauts{14}" : Bool = PLC Défauts.Defauts[14] AT %DB13.DBX1.6, 1 s
   "Défauts_Defauts{15}" : Bool = PLC Défauts.Defauts[15] AT %DB13.DBX1.7, 1 s
   "Défauts_Defauts{3}" : Bool = PLC Défauts.Defauts[3] AT %DB13.DBX0.3, 1 s
   "Défauts_Defauts{4}" : Bool = PLC Défauts.Defauts[4] AT %DB13.DBX0.4, 1 s
   "Défauts_Defauts{5}" : Bool = PLC Défauts.Defauts[5] AT %DB13.DBX0.5, 1 s
   "Défauts_Defauts{6}" : Bool = PLC Défauts.Defauts[6] AT %DB13.DBX0.6, 1 s
   "Défauts_Defauts{7}" : Bool = PLC Défauts.Defauts[7] AT %DB13.DBX0.7, 1 s
   "Défauts_Defauts{8}" : Bool = PLC Défauts.Defauts[8] AT %DB13.DBX1.0, 1 s
   "Défauts_Defauts{9}" : Bool = PLC Défauts.Defauts[9] AT %DB13.DBX1.1, 1 s
   "Défauts_Defauts{10}" : Bool = PLC Défauts.Defauts[10] AT %DB13.DBX1.2, 1 s
   "Défauts_Defauts{11}" : Bool = PLC Défauts.Defauts[11] AT %DB13.DBX1.3, 1 s
   "Défauts_Defauts{16}" : Bool = PLC Défauts.Defauts[16] AT %DB13.DBX2.0, 1 s
   "Défauts_Defauts{17}" : Bool = PLC Défauts.Defauts[17] AT %DB13.DBX2.1, 1 s
   "Défauts_Defauts{20}" : Bool = PLC Défauts.Defauts[20] AT %DB13.DBX2.4, 1 s
   "Défauts_Defauts{21}" : Bool = PLC Défauts.Defauts[21] AT %DB13.DBX2.5, 1 s
   "Défauts_Defauts{22}" : Bool = PLC Défauts.Defauts[22] AT %DB13.DBX2.6, 1 s
   "Défauts_Defauts{23}" : Bool = PLC Défauts.Defauts[23] AT %DB13.DBX2.7, 1 s
   "Défauts_Defauts{24}" : Bool = PLC Défauts.Defauts[24] AT %DB13.DBX3.0, 1 s
   "Défauts_Defauts{25}" : Bool = PLC Défauts.Defauts[25] AT %DB13.DBX3.1, 1 s
   "Défauts_Defauts{26}" : Bool = PLC Défauts.Defauts[26] AT %DB13.DBX3.2, 1 s
   "Q_Wieland_Acces_Autorisé" : Bool = PLC Q_Wieland_Acces_Autorisé AT %Q18.0, 1 s
   "I_Wieland_Au_armoire" : Bool = PLC I_Wieland_Au_armoire AT %I16.0, 1 s
   "I_Wieland_Au_porte01" : Bool = PLC I_Wieland_Au_porte01 AT %I16.1, 1 s
   "I_Wieland_Au_Porte02" : Bool = PLC I_Wieland_Au_Porte02 AT %I16.2, 1 s
   "I_Wieland_Au_Robot01_Fanuc" : Bool = PLC I_Wieland_Au_Robot01_Fanuc AT %I16.3, 1 s
   "I_Wieland_Au_Robot02_Fanuc" : Bool = PLC I_Wieland_Au_Robot02_Fanuc AT %I16.4, 1 s
   "I_Wieland_Au_Robot03_ABB" : Bool = PLC I_Wieland_Au_Robot03_ABB AT %I16.5, 1 s
   "I_Wielmand_Au_Robot04_UR" : Bool = PLC I_Wielmand_Au_Robot04_UR AT %I16.6, 1 s
   "I_Wieland_Au_Robot05_UR" : Bool = PLC I_Wieland_Au_Robot05_UR AT %I16.7, 1 s
   "I_wieland_Au_Carroussel" : Bool = PLC I_wieland_Au_Carroussel AT %I17.0, 1 s
   "I_Wieland_Au_Carterisation" : Bool = PLC I_Wieland_Au_Carterisation AT %I17.1, 1 s
   "I_Wieland_Rearmement" : Bool = PLC I_Wieland_Rearmement AT %I17.4, 1 s
   "I_Wieland_Dmd acces" : Bool = PLC "I_Wieland_Dmd acces" AT %I17.5, 1 s
   "I_Wieland_Mise sous puissance" : Bool = PLC "I_Wieland_Mise sous puissance" AT %I17.6, 1 s
   "I_Wieland_Mise hors puissance" : Bool = PLC "I_Wieland_Mise hors puissance" AT %I17.7, 1 s
   "I_Wieland_Acces_autorisé" : Bool = PLC I_Wieland_Acces_autorisé AT %I18.0, 1 s
   "I_Wieland_rearmement_Porte" : Bool = PLC I_Wieland_rearmement_Porte AT %I18.1, 1 s
   "I_Wieland_En_Service" : Bool = PLC I_Wieland_En_Service AT %I18.2, 1 s
   "I_Wieland_Porte_non_Réarmée" : Bool = PLC I_Wieland_Porte_non_Réarmée AT %I18.3, 1 s
   "I_porte_vision_op" : Bool = PLC I_porte_vision_op AT %I7.6, 1 s
   "I_porte_vision_cl" : Bool = PLC I_porte_vision_cl AT %I6.6, 1 s
   "Var_Convoyeur_Carton_ConvoyeurC01_Reserve01" : Bool = PLC DB_Variateurs.ConvoyeurC01.Cmd.Reserve01 AT %DB17.DBX4.0, 1 s
   "Var_Convoyeur_Carton_ConvoyeurC01_Reserve02" : Bool = PLC DB_Variateurs.ConvoyeurC01.Cmd.Reserve02 AT %DB17.DBX4.1, 1 s
   "Var_Convoyeur_Carton_ConvoyeurC01_PilotageParApi" : Bool = PLC DB_Variateurs.ConvoyeurC01.Cmd.PilotageParApi AT %DB17.DBX4.2, 1 s
   "Var_Convoyeur_Carton_ConvoyeurC01_InversionConsigne" : Bool = PLC DB_Variateurs.ConvoyeurC01.Cmd.InversionConsigne AT %DB17.DBX4.3, 1 s
   "Var_Convoyeur_Carton_ConvoyeurC01_Reserve03" : Bool = PLC DB_Variateurs.ConvoyeurC01.Cmd.Reserve03 AT %DB17.DBX4.4, 1 s
   "Var_Convoyeur_Carton_ConvoyeurC01_PotPlus" : Bool = PLC DB_Variateurs.ConvoyeurC01.Cmd.PotPlus AT %DB17.DBX4.5, 1 s
   "Var_Convoyeur_Carton_ConvoyeurC01_PotMoins" : Bool = PLC DB_Variateurs.ConvoyeurC01.Cmd.PotMoins AT %DB17.DBX4.6, 1 s
   "Var_Convoyeur_Carton_ConvoyeurC01_Reserve04" : Bool = PLC DB_Variateurs.ConvoyeurC01.Cmd.Reserve04 AT %DB17.DBX4.7, 1 s
   "Var_Convoyeur_Carton_ConvoyeurC01_Marche" : Bool = PLC DB_Variateurs.ConvoyeurC01.Cmd.Marche AT %DB17.DBX5.0, 1 s
   "Var_Convoyeur_Carton_ConvoyeurC01_Arret2" : Bool = PLC DB_Variateurs.ConvoyeurC01.Cmd.Arret2 AT %DB17.DBX5.1, 1 s
   "Var_Convoyeur_Carton_ConvoyeurC01_Arret3" : Bool = PLC DB_Variateurs.ConvoyeurC01.Cmd.Arret3 AT %DB17.DBX5.2, 1 s
   "Var_Convoyeur_Carton_ConvoyeurC01_DebloqFonctionnement" : Bool = PLC DB_Variateurs.ConvoyeurC01.Cmd.DebloqFonctionnement AT %DB17.DBX5.3, 1 s
   "Var_Convoyeur_Carton_ConvoyeurC01_DebloqRampe" : Bool = PLC DB_Variateurs.ConvoyeurC01.Cmd.DebloqRampe AT %DB17.DBX5.4, 1 s
   "Var_Convoyeur_Carton_ConvoyeurC01_GelerGenerateurRampe" : Bool = PLC DB_Variateurs.ConvoyeurC01.Cmd.GelerGenerateurRampe AT %DB17.DBX5.5, 1 s
   "Var_Convoyeur_Carton_ConvoyeurC01_DebloqConsigne" : Bool = PLC DB_Variateurs.ConvoyeurC01.Cmd.DebloqConsigne AT %DB17.DBX5.6, 1 s
   "Var_Convoyeur_Carton_ConvoyeurC01_AcquitDefaut" : Bool = PLC DB_Variateurs.ConvoyeurC01.Cmd.AcquitDefaut AT %DB17.DBX5.7, 1 s
   "Var_Convoyeur_Carton_ConvoyeurC01_Consigne" : Int = PLC DB_Variateurs.ConvoyeurC01.Cmd.Consigne AT %DB17.DBW6, 1 s
   "Var_Convoyeur_Carton_ConvoyeurC01_EcartVitesse" : Bool = PLC DB_Variateurs.ConvoyeurC01.Status.EcartVitesse AT %DB17.DBX0.0, 1 s
   "Var_Convoyeur_Carton_ConvoyeurC01_CommandeDemander" : Bool = PLC DB_Variateurs.ConvoyeurC01.Status.CommandeDemander AT %DB17.DBX0.1, 1 s
   "Var_Convoyeur_Carton_ConvoyeurC01_VitesseMaxAtteinte" : Bool = PLC DB_Variateurs.ConvoyeurC01.Status.VitesseMaxAtteinte AT %DB17.DBX0.2, 1 s
   "Var_Convoyeur_Carton_ConvoyeurC01_Limite" : Bool = PLC DB_Variateurs.ConvoyeurC01.Status.Limite AT %DB17.DBX0.3, 1 s
   "Var_Convoyeur_Carton_ConvoyeurC01_FreinMoteur" : Bool = PLC DB_Variateurs.ConvoyeurC01.Status.FreinMoteur AT %DB17.DBX0.4, 1 s
   "Var_Convoyeur_Carton_ConvoyeurC01_AlarmeSurchauffe" : Bool = PLC DB_Variateurs.ConvoyeurC01.Status.AlarmeSurchauffe AT %DB17.DBX0.5, 1 s
   "Var_Convoyeur_Carton_ConvoyeurC01_MoteurSensAvant" : Bool = PLC DB_Variateurs.ConvoyeurC01.Status.MoteurSensAvant AT %DB17.DBX0.6, 1 s
   "Var_Convoyeur_Carton_ConvoyeurC01_SurchargeMoteur" : Bool = PLC DB_Variateurs.ConvoyeurC01.Status.SurchargeMoteur AT %DB17.DBX0.7, 1 s
   "Var_Convoyeur_Carton_ConvoyeurC01_PretEnclenchement" : Bool = PLC DB_Variateurs.ConvoyeurC01.Status.PretEnclenchement AT %DB17.DBX1.0, 1 s
   "Var_Convoyeur_Carton_ConvoyeurC01_PretFonctionnement" : Bool = PLC DB_Variateurs.ConvoyeurC01.Status.PretFonctionnement AT %DB17.DBX1.1, 1 s
   "Var_Convoyeur_Carton_ConvoyeurC01_Fonctionnement_Debloq" : Bool = PLC DB_Variateurs.ConvoyeurC01.Status.Fonctionnement_Debloq AT %DB17.DBX1.2, 1 s
   "Var_Convoyeur_Carton_ConvoyeurC01_DefautActif" : Bool = PLC DB_Variateurs.ConvoyeurC01.Status.DefautActif AT %DB17.DBX1.3, 1 s
   "Var_Convoyeur_Carton_ConvoyeurC01_Arret2Etat" : Bool = PLC DB_Variateurs.ConvoyeurC01.Status.Arret2Etat AT %DB17.DBX1.4, 1 s
   "Var_Convoyeur_Carton_ConvoyeurC01_Arret3Etat" : Bool = PLC DB_Variateurs.ConvoyeurC01.Status.Arret3Etat AT %DB17.DBX1.5, 1 s
   "Var_Convoyeur_Carton_ConvoyeurC01_BlocageActif" : Bool = PLC DB_Variateurs.ConvoyeurC01.Status.BlocageActif AT %DB17.DBX1.6, 1 s
   "Var_Convoyeur_Carton_ConvoyeurC01_AlarmeActive" : Bool = PLC DB_Variateurs.ConvoyeurC01.Status.AlarmeActive AT %DB17.DBX1.7, 1 s
   "Var_Convoyeur_Carton_ConvoyeurC01_Vitesse" : Int = PLC DB_Variateurs.ConvoyeurC01.Status.Vitesse AT %DB17.DBW2, 1 s
   "Var_Convoyeur_Carton_ConvoyeurC02_Reserve01" : Bool = PLC DB_Variateurs.ConvoyeurC02.Cmd.Reserve01 AT %DB17.DBX12.0, 1 s
   "Var_Convoyeur_Carton_ConvoyeurC02_Reserve02" : Bool = PLC DB_Variateurs.ConvoyeurC02.Cmd.Reserve02 AT %DB17.DBX12.1, 1 s
   "Var_Convoyeur_Carton_ConvoyeurC02_PilotageParApi" : Bool = PLC DB_Variateurs.ConvoyeurC02.Cmd.PilotageParApi AT %DB17.DBX12.2, 1 s
   "Var_Convoyeur_Carton_ConvoyeurC02_InversionConsigne" : Bool = PLC DB_Variateurs.ConvoyeurC02.Cmd.InversionConsigne AT %DB17.DBX12.3, 1 s
   "Var_Convoyeur_Carton_ConvoyeurC02_Reserve03" : Bool = PLC DB_Variateurs.ConvoyeurC02.Cmd.Reserve03 AT %DB17.DBX12.4, 1 s
   "Var_Convoyeur_Carton_ConvoyeurC02_PotPlus" : Bool = PLC DB_Variateurs.ConvoyeurC02.Cmd.PotPlus AT %DB17.DBX12.5, 1 s
   "Var_Convoyeur_Carton_ConvoyeurC02_PotMoins" : Bool = PLC DB_Variateurs.ConvoyeurC02.Cmd.PotMoins AT %DB17.DBX12.6, 1 s
   "Var_Convoyeur_Carton_ConvoyeurC02_Reserve04" : Bool = PLC DB_Variateurs.ConvoyeurC02.Cmd.Reserve04 AT %DB17.DBX12.7, 1 s
   "Var_Convoyeur_Carton_ConvoyeurC02_Marche" : Bool = PLC DB_Variateurs.ConvoyeurC02.Cmd.Marche AT %DB17.DBX13.0, 1 s
   "Var_Convoyeur_Carton_ConvoyeurC02_Arret2" : Bool = PLC DB_Variateurs.ConvoyeurC02.Cmd.Arret2 AT %DB17.DBX13.1, 1 s
   "Var_Convoyeur_Carton_ConvoyeurC02_Arret3" : Bool = PLC DB_Variateurs.ConvoyeurC02.Cmd.Arret3 AT %DB17.DBX13.2, 1 s
   "Var_Convoyeur_Carton_ConvoyeurC02_DebloqFonctionnement" : Bool = PLC DB_Variateurs.ConvoyeurC02.Cmd.DebloqFonctionnement AT %DB17.DBX13.3, 1 s
   "Var_Convoyeur_Carton_ConvoyeurC02_DebloqRampe" : Bool = PLC DB_Variateurs.ConvoyeurC02.Cmd.DebloqRampe AT %DB17.DBX13.4, 1 s
   "Var_Convoyeur_Carton_ConvoyeurC02_GelerGenerateurRampe" : Bool = PLC DB_Variateurs.ConvoyeurC02.Cmd.GelerGenerateurRampe AT %DB17.DBX13.5, 1 s
   "Var_Convoyeur_Carton_ConvoyeurC02_DebloqConsigne" : Bool = PLC DB_Variateurs.ConvoyeurC02.Cmd.DebloqConsigne AT %DB17.DBX13.6, 1 s
   "Var_Convoyeur_Carton_ConvoyeurC02_AcquitDefaut" : Bool = PLC DB_Variateurs.ConvoyeurC02.Cmd.AcquitDefaut AT %DB17.DBX13.7, 1 s
   "Var_Convoyeur_Carton_ConvoyeurC02_Consigne" : Int = PLC DB_Variateurs.ConvoyeurC02.Cmd.Consigne AT %DB17.DBW14, 1 s
   "Var_Convoyeur_Carton_ConvoyeurC02_EcartVitesse" : Bool = PLC DB_Variateurs.ConvoyeurC02.Status.EcartVitesse AT %DB17.DBX8.0, 1 s
   "Var_Convoyeur_Carton_ConvoyeurC02_CommandeDemander" : Bool = PLC DB_Variateurs.ConvoyeurC02.Status.CommandeDemander AT %DB17.DBX8.1, 1 s
   "Var_Convoyeur_Carton_ConvoyeurC02_VitesseMaxAtteinte" : Bool = PLC DB_Variateurs.ConvoyeurC02.Status.VitesseMaxAtteinte AT %DB17.DBX8.2, 1 s
   "Var_Convoyeur_Carton_ConvoyeurC02_Limite" : Bool = PLC DB_Variateurs.ConvoyeurC02.Status.Limite AT %DB17.DBX8.3, 1 s
   "Var_Convoyeur_Carton_ConvoyeurC02_FreinMoteur" : Bool = PLC DB_Variateurs.ConvoyeurC02.Status.FreinMoteur AT %DB17.DBX8.4, 1 s
   "Var_Convoyeur_Carton_ConvoyeurC02_AlarmeSurchauffe" : Bool = PLC DB_Variateurs.ConvoyeurC02.Status.AlarmeSurchauffe AT %DB17.DBX8.5, 1 s
   "Var_Convoyeur_Carton_ConvoyeurC02_MoteurSensAvant" : Bool = PLC DB_Variateurs.ConvoyeurC02.Status.MoteurSensAvant AT %DB17.DBX8.6, 1 s
   "Var_Convoyeur_Carton_ConvoyeurC02_SurchargeMoteur" : Bool = PLC DB_Variateurs.ConvoyeurC02.Status.SurchargeMoteur AT %DB17.DBX8.7, 1 s
   "Var_Convoyeur_Carton_ConvoyeurC02_PretEnclenchement" : Bool = PLC DB_Variateurs.ConvoyeurC02.Status.PretEnclenchement AT %DB17.DBX9.0, 1 s
   "Var_Convoyeur_Carton_ConvoyeurC02_PretFonctionnement" : Bool = PLC DB_Variateurs.ConvoyeurC02.Status.PretFonctionnement AT %DB17.DBX9.1, 1 s
   "Var_Convoyeur_Carton_ConvoyeurC02_Fonctionnement_Debloq" : Bool = PLC DB_Variateurs.ConvoyeurC02.Status.Fonctionnement_Debloq AT %DB17.DBX9.2, 1 s
   "Var_Convoyeur_Carton_ConvoyeurC02_DefautActif" : Bool = PLC DB_Variateurs.ConvoyeurC02.Status.DefautActif AT %DB17.DBX9.3, 1 s
   "Var_Convoyeur_Carton_ConvoyeurC02_Arret2Etat" : Bool = PLC DB_Variateurs.ConvoyeurC02.Status.Arret2Etat AT %DB17.DBX9.4, 1 s
   "Var_Convoyeur_Carton_ConvoyeurC02_Arret3Etat" : Bool = PLC DB_Variateurs.ConvoyeurC02.Status.Arret3Etat AT %DB17.DBX9.5, 1 s
   "Var_Convoyeur_Carton_ConvoyeurC02_BlocageActif" : Bool = PLC DB_Variateurs.ConvoyeurC02.Status.BlocageActif AT %DB17.DBX9.6, 1 s
   "Var_Convoyeur_Carton_ConvoyeurC02_AlarmeActive" : Bool = PLC DB_Variateurs.ConvoyeurC02.Status.AlarmeActive AT %DB17.DBX9.7, 1 s
   "Var_Convoyeur_Carton_ConvoyeurC02_Vitesse" : Int = PLC DB_Variateurs.ConvoyeurC02.Status.Vitesse AT %DB17.DBW10, 1 s
   "Var_Convoyeur_Carton_ConvoyeurC03_Reserve01" : Bool = PLC DB_Variateurs.ConvoyeurC03.Cmd.Reserve01 AT %DB17.DBX20.0, 1 s
   "Var_Convoyeur_Carton_ConvoyeurC03_Reserve02" : Bool = PLC DB_Variateurs.ConvoyeurC03.Cmd.Reserve02 AT %DB17.DBX20.1, 1 s
   "Var_Convoyeur_Carton_ConvoyeurC03_PilotageParApi" : Bool = PLC DB_Variateurs.ConvoyeurC03.Cmd.PilotageParApi AT %DB17.DBX20.2, 1 s
   "Var_Convoyeur_Carton_ConvoyeurC03_InversionConsigne" : Bool = PLC DB_Variateurs.ConvoyeurC03.Cmd.InversionConsigne AT %DB17.DBX20.3, 1 s
   "Var_Convoyeur_Carton_ConvoyeurC03_Reserve03" : Bool = PLC DB_Variateurs.ConvoyeurC03.Cmd.Reserve03 AT %DB17.DBX20.4, 1 s
   "Var_Convoyeur_Carton_ConvoyeurC03_PotPlus" : Bool = PLC DB_Variateurs.ConvoyeurC03.Cmd.PotPlus AT %DB17.DBX20.5, 1 s
   "Var_Convoyeur_Carton_ConvoyeurC03_PotMoins" : Bool = PLC DB_Variateurs.ConvoyeurC03.Cmd.PotMoins AT %DB17.DBX20.6, 1 s
   "Var_Convoyeur_Carton_ConvoyeurC03_Reserve04" : Bool = PLC DB_Variateurs.ConvoyeurC03.Cmd.Reserve04 AT %DB17.DBX20.7, 1 s
   "Var_Convoyeur_Carton_ConvoyeurC03_Marche" : Bool = PLC DB_Variateurs.ConvoyeurC03.Cmd.Marche AT %DB17.DBX21.0, 1 s
   "Var_Convoyeur_Carton_ConvoyeurC03_Arret2" : Bool = PLC DB_Variateurs.ConvoyeurC03.Cmd.Arret2 AT %DB17.DBX21.1, 1 s
   "Var_Convoyeur_Carton_ConvoyeurC03_Arret3" : Bool = PLC DB_Variateurs.ConvoyeurC03.Cmd.Arret3 AT %DB17.DBX21.2, 1 s
   "Var_Convoyeur_Carton_ConvoyeurC03_DebloqFonctionnement" : Bool = PLC DB_Variateurs.ConvoyeurC03.Cmd.DebloqFonctionnement AT %DB17.DBX21.3, 1 s
   "Var_Convoyeur_Carton_ConvoyeurC03_DebloqRampe" : Bool = PLC DB_Variateurs.ConvoyeurC03.Cmd.DebloqRampe AT %DB17.DBX21.4, 1 s
   "Var_Convoyeur_Carton_ConvoyeurC03_GelerGenerateurRampe" : Bool = PLC DB_Variateurs.ConvoyeurC03.Cmd.GelerGenerateurRampe AT %DB17.DBX21.5, 1 s
   "Var_Convoyeur_Carton_ConvoyeurC03_DebloqConsigne" : Bool = PLC DB_Variateurs.ConvoyeurC03.Cmd.DebloqConsigne AT %DB17.DBX21.6, 1 s
   "Var_Convoyeur_Carton_ConvoyeurC03_AcquitDefaut" : Bool = PLC DB_Variateurs.ConvoyeurC03.Cmd.AcquitDefaut AT %DB17.DBX21.7, 1 s
   "Var_Convoyeur_Carton_ConvoyeurC03_Consigne" : Int = PLC DB_Variateurs.ConvoyeurC03.Cmd.Consigne AT %DB17.DBW22, 1 s
   "Var_Convoyeur_Carton_ConvoyeurC03_EcartVitesse" : Bool = PLC DB_Variateurs.ConvoyeurC03.Status.EcartVitesse AT %DB17.DBX16.0, 1 s
   "Var_Convoyeur_Carton_ConvoyeurC03_CommandeDemander" : Bool = PLC DB_Variateurs.ConvoyeurC03.Status.CommandeDemander AT %DB17.DBX16.1, 1 s
   "Var_Convoyeur_Carton_ConvoyeurC03_VitesseMaxAtteinte" : Bool = PLC DB_Variateurs.ConvoyeurC03.Status.VitesseMaxAtteinte AT %DB17.DBX16.2, 1 s
   "Var_Convoyeur_Carton_ConvoyeurC03_Limite" : Bool = PLC DB_Variateurs.ConvoyeurC03.Status.Limite AT %DB17.DBX16.3, 1 s
   "Var_Convoyeur_Carton_ConvoyeurC03_FreinMoteur" : Bool = PLC DB_Variateurs.ConvoyeurC03.Status.FreinMoteur AT %DB17.DBX16.4, 1 s
   "Var_Convoyeur_Carton_ConvoyeurC03_AlarmeSurchauffe" : Bool = PLC DB_Variateurs.ConvoyeurC03.Status.AlarmeSurchauffe AT %DB17.DBX16.5, 1 s
   "Var_Convoyeur_Carton_ConvoyeurC03_MoteurSensAvant" : Bool = PLC DB_Variateurs.ConvoyeurC03.Status.MoteurSensAvant AT %DB17.DBX16.6, 1 s
   "Var_Convoyeur_Carton_ConvoyeurC03_SurchargeMoteur" : Bool = PLC DB_Variateurs.ConvoyeurC03.Status.SurchargeMoteur AT %DB17.DBX16.7, 1 s
   "Var_Convoyeur_Carton_ConvoyeurC03_PretEnclenchement" : Bool = PLC DB_Variateurs.ConvoyeurC03.Status.PretEnclenchement AT %DB17.DBX17.0, 1 s
   "Var_Convoyeur_Carton_ConvoyeurC03_PretFonctionnement" : Bool = PLC DB_Variateurs.ConvoyeurC03.Status.PretFonctionnement AT %DB17.DBX17.1, 1 s
   "Var_Convoyeur_Carton_ConvoyeurC03_Fonctionnement_Debloq" : Bool = PLC DB_Variateurs.ConvoyeurC03.Status.Fonctionnement_Debloq AT %DB17.DBX17.2, 1 s
   "Var_Convoyeur_Carton_ConvoyeurC03_DefautActif" : Bool = PLC DB_Variateurs.ConvoyeurC03.Status.DefautActif AT %DB17.DBX17.3, 1 s
   "Var_Convoyeur_Carton_ConvoyeurC03_Arret2Etat" : Bool = PLC DB_Variateurs.ConvoyeurC03.Status.Arret2Etat AT %DB17.DBX17.4, 1 s
   "Var_Convoyeur_Carton_ConvoyeurC03_Arret3Etat" : Bool = PLC DB_Variateurs.ConvoyeurC03.Status.Arret3Etat AT %DB17.DBX17.5, 1 s
   "Var_Convoyeur_Carton_ConvoyeurC03_BlocageActif" : Bool = PLC DB_Variateurs.ConvoyeurC03.Status.BlocageActif AT %DB17.DBX17.6, 1 s
   "Var_Convoyeur_Carton_ConvoyeurC03_AlarmeActive" : Bool = PLC DB_Variateurs.ConvoyeurC03.Status.AlarmeActive AT %DB17.DBX17.7, 1 s
   "Var_Convoyeur_Carton_ConvoyeurC03_Vitesse" : Int = PLC DB_Variateurs.ConvoyeurC03.Status.Vitesse AT %DB17.DBW18, 1 s
   "Parametres_Sp_vitesse_manu_C01" : Int = PLC Parametres.Convoyeurs.Manu.i_Vitesse_manu_C01, 1 s
   "Parametres_Sp_vitesse_manu_C02" : Int = PLC Parametres.Convoyeurs.Manu.i_Vitesse_manu_C02, 1 s
   "Parametres_Sp_vitesse_manu_C03" : Int = PLC Parametres.Convoyeurs.Manu.i_Vitesse_manu_C03, 1 s
   "I_Wieland_Porte 01 ouverte" : Bool = PLC "I_Wieland_Porte 01 ouverte" AT %I17.2, 1 s
   "I_Wieland_Porte 02 Ouverte" : Bool = PLC "I_Wieland_Porte 02 Ouverte" AT %I17.3, 1 s
   "Touche_Tch_Manu{90}" : Bool = PLC Tch_HMI.Tch_Manu[90], 1 s
   "Touche_Tch_Manu{91}" : Bool = PLC Tch_HMI.Tch_Manu[91], 1 s
   "Bits_B_init_cours" : Bool = PLC Bits_Globaux.x_Init_en_cours, 1 s
   "Bits_B_dmd_Init_robot" : Bool = PLC Bits_Globaux.x_Dmd_Init_robot, 1 s
   "B_Pret_TP_Robotique" : Bool = PLC Voyants_HMI.x_VOY_Tp_robot_pret AT %DB1.DBX0.0, 500 ms
   "Fanuc1_Auto" : Bool = PLC Fanuc01_Selecteur_Auto AT %I30.4, 1 s
   "Fanuc2_Auto" : Bool = PLC Fanuc02_Selecteur_Auto AT %I220.4, 1 s
   "Fanuc1_Autor_Prise" : Bool = PLC Fanuc01_Autor_Prise AT %Q40.5, 1 s
   "Fanuc2_Autor_Prise" : Bool = PLC Fanuc02_Autor_Prise AT %Q31.5, 1 s
   "Fanuc2_Autor_Depose" : Bool = PLC Fanuc02_Autor_Depose AT %Q31.6, 1 s
   "Fanuc1_Autor_vers_Fanuc02" : Bool = PLC Fanuc01_envoi_signal_pret_vers_fanuc02 AT %Q31.7, 1 s
   "Robots_En_Auto" : Bool = PLC Bits_Globaux.x_Robots_en_AUTO AT %M200.0, 1 s
   "Défauts_Def_Canal03" : Int = PLC Défauts.Def_Canal03 AT %DB13.DBW18, 1 s
   "Bits_Pret_Demo_Hippo" : Bool = PLC Voyants_HMI.x_VOY_Demo_pret, 500 ms
   "Bits_B_TP_Robot" : Bool = PLC Tch_HMI.Tch_Tp_Robot, 500 ms
   "B_VOY_DCY" : Bool = PLC Voyants_HMI.x_VOY_DCY, 500 ms
   "B_VOY_ACY" : Bool = PLC Voyants_HMI.x_VOY_ACY, 500 ms
   "VOY_Init" : Bool = PLC Voyants_HMI.x_VOY_INIT, 1 s
   "Bits_Init_glob_OK" : Bool = PLC Bits_Globaux.x_Init_glob_OK, 1 s
   "FanucR1_In_auto" : Bool = PLC Fanuc_R1_DB.DATA.status.x_In_auto_mode, 1 s
   "FanucR2_In_Auto" : Bool = PLC Fanuc_R2_DB.DATA.status.x_In_auto_mode, 1 s
   "Fanuc1_Teach_active" : Bool = PLC Fanuc_R1_DB.DATA.status.x_Teach_on, 1 s
   "Fanuc2_teach_active" : Bool = PLC Fanuc_R2_DB.DATA.status.x_Teach_on, 1 s
   "CV01_Hipp_Marche" : Bool = PLC DB_Convoyeurs_Hipp.Convoyeur[1].Status.x_EnMarche, 1 s
   "CV03_Hipp_Marche" : Bool = PLC DB_Convoyeurs_Hipp.Convoyeur[3].Status.x_EnMarche, 1 s
   "CV02_Hipp_Marche" : Bool = PLC DB_Convoyeurs_Hipp.Convoyeur[2].Status.x_EnMarche, 1 s
   "CV04_Hipp_Marche" : Bool = PLC DB_Convoyeurs_Hipp.Convoyeur[4].Status.x_EnMarche, 1 s
   "Touche_Tch_Manu{92}" : Bool = PLC Tch_HMI.Tch_Manu[92], 1 s   // Envoi trigger Vision Keyence
   "Touche_Tch_Manu{93}" : Bool = PLC Tch_HMI.Tch_Manu[93], 1 s   // Envoi trigger Vision Keyence
   "Touche_Tch_Manu{94}" : Bool = PLC Tch_HMI.Tch_Manu[94], 1 s
   "Touche_Tch_Manu{95}" : Bool = PLC Tch_HMI.Tch_Manu[95], 1 s
   "Touche_Tch_Manu{96}" : Bool = PLC Tch_HMI.Tch_Manu[96], 1 s

HMI tags "DB_Stations"
   "DB_Stations_Station{1}" : Station_Hipp = PLC DB_Stations.Station[1], 1 s
   "DB_Stations_Station{2}" : Station_Hipp = PLC DB_Stations.Station[2], 1 s
   "DB_Stations_Station{3}" : Station_Hipp = PLC DB_Stations.Station[3], 1 s
   "DB_Stations_Station{4}" : Station_Hipp = PLC DB_Stations.Station[4], 1 s
   "DB_Stations_Station{5}" : Station_Hipp = PLC DB_Stations.Station[5], 1 s
   "DB_Stations_Station{6}" : Station_Hipp = PLC DB_Stations.Station[6], 1 s
   "DB_Stations_Station{7}" : Station_Hipp = PLC DB_Stations.Station[7], 1 s

HMI tags "Bits_generaux"
   "Bits_Globaux_x_Init_glob_OK" : Bool = PLC Bits_Globaux.x_Init_glob_OK, 1 s
   "Bits_Globaux_x_Defaut_non_bloquant" : Bool = PLC Bits_Globaux.x_Defaut_non_bloquant, 1 s
   "Bits_Globaux_x_Demo_Hippo_en_cours" : Bool = PLC Bits_Globaux.x_Demo_Hippo_en_cours, 1 s
   "Bits_Globaux_x_En_service" : Bool = PLC Bits_Globaux.x_En_service, 1 s
   "Bits_Globaux_x_En_auto" : Bool = PLC Bits_Globaux.x_En_auto, 1 s
   "Bits_Globaux_x_En_manu" : Bool = PLC Bits_Globaux.x_En_manu, 1 s
   "Bits_Globaux_x_Dmd_Init_robot" : Bool = PLC Bits_Globaux.x_Dmd_Init_robot, 1 s
   "Bits_Globaux_x_Init_en_cours" : Bool = PLC Bits_Globaux.x_Init_en_cours, 1 s
   "Bits_Globaux_x_Defaut_bloquant" : Bool = PLC Bits_Globaux.x_Defaut_bloquant, 1 s
   "Bits_Globaux_x_Robots_en_AUTO" : Bool = PLC Bits_Globaux.x_Robots_en_AUTO, 1 s
   "Bits_Globaux_x_Tp_Robots_en_cours" : Bool = PLC Bits_Globaux.x_Tp_Robots_en_cours, 1 s
   "Bits_Globaux_x_En_cycle_auto" : Bool = PLC Bits_Globaux.x_En_cycle_auto AT %DB1.DBX0.0, 1 s

HMI tags "VoyantsHMI"
   "Voyants_HMI_x_VOY_Demo_pret" : Bool = PLC Voyants_HMI.x_VOY_Demo_pret, 500 ms
   "Voyants_HMI_x_VOY_Tp_robot_pret" : Bool = PLC Voyants_HMI.x_VOY_Tp_robot_pret, 500 ms
   "Voyants_HMI_x_VOY_DCY" : Bool = PLC Voyants_HMI.x_VOY_DCY, 500 ms
   "Voyants_HMI_x_VOY_ACY" : Bool = PLC Voyants_HMI.x_VOY_ACY, 500 ms
   "Voyants_HMI_x_VOY_INIT" : Bool = PLC Voyants_HMI.x_VOY_INIT, 500 ms
   "Voyants_HMI_x_VOY_Init_requis_en_auto" : Bool = PLC Voyants_HMI.x_VOY_Init_requis_en_auto, 500 ms

HMI tags "DB_Imprimantes"
   "DB_Imprimantes_Imprimante{1}" : Imprimante3D = PLC DB_Imprimantes.Imprimante[1], 1 s
   "DB_Imprimantes_Imprimante{2}" : Imprimante3D = PLC DB_Imprimantes.Imprimante[2], 1 s
   "DB_Imprimantes_Imprimante{3}" : Imprimante3D = PLC DB_Imprimantes.Imprimante[3], 1 s
   "DB_Imprimantes_Imprimante{4}" : Imprimante3D = PLC DB_Imprimantes.Imprimante[4], 1 s

HMI tags "DB_UR4"
   "40_UR_R4_DB_DATA" : UR_Cobot = PLC "40_UR_R4_DB".DATA, 1 s

HMI tags "DB_UR5"
   "60_UR_R5_DB_DATA" : UR_Cobot = PLC "60_UR_R5_DB".DATA, 1 s

HMI tags "DB_porte_vision"
   "32_Cmd_porte_vision_DB_x_ouverture_porte_vision" : Bool = PLC "32_Cmd_porte_vision_DB".x_ouverture_porte_vision, 1 s
   "32_Cmd_porte_vision_DB_x_fermeture_porte_vision" : Bool = PLC "32_Cmd_porte_vision_DB".x_fermeture_porte_vision, 1 s
   "32_Cmd_porte_vision_DB_x_Ouverture_porte_manu" : Bool = PLC "32_Cmd_porte_vision_DB".x_Ouverture_porte_manu, 1 s
   "32_Cmd_porte_vision_DB_x_Fermeture_porte_manu" : Bool = PLC "32_Cmd_porte_vision_DB".x_Fermeture_porte_manu, 1 s

discrete alarms
   1: 'Défaut verin de blocage 01', class Errors, trigger "Défauts_Def_Canal01" bit 8
   2: 'Défaut verin de blocage 02', class Errors, trigger "Défauts_Def_Canal01" bit 9
   3: 'Défaut verin de blocage 03', class Errors, trigger "Défauts_Def_Canal01" bit 10
   4: 'Défaut verin de blocage 04', class Errors, trigger "Défauts_Def_Canal01" bit 11
   5: 'Défaut elevateur 01', class Errors, trigger "Défauts_Def_Canal01" bit 12
   6: 'Défaut elevateur 02', class Errors, trigger "Défauts_Def_Canal01" bit 13
   7: 'Défaut elevateur 03', class Errors, trigger "Défauts_Def_Canal01" bit 14
   8: 'Défaut elevateur 04', class Errors, trigger "Défauts_Def_Canal01" bit 15
   9: 'Défaut elevateur 05', class Errors, trigger "Défauts_Def_Canal01" bit 0
   10: 'Défaut elevateur 06', class Errors, trigger "Défauts_Def_Canal01" bit 1
   11: 'Défaut elevateur 07', class Errors, trigger "Défauts_Def_Canal01" bit 2
   12: 'Défaut Convoyeur hyppodrome 01', class Errors, trigger "Défauts_Def_Canal01" bit 3
   13: 'Défaut Convoyeur hyppodrome 02', class Errors, trigger "Défauts_Def_Canal01" bit 4
   14: 'Défaut Convoyeur hyppodrome 03', class Errors, trigger "Défauts_Def_Canal01" bit 5
   15: 'Défaut Convoyeur hyppodrome 04', class Errors, trigger "Défauts_Def_Canal01" bit 6
   16: 'Défaut Convoyeur Carton 01', class Errors, trigger "Défauts_Def_Canal01" bit 7
   17: 'Défaut Convoyeur Carton 02', class Errors, trigger "Défauts_Def_Canal02" bit 8
   18: 'Défaut Convoyeur Carton 03', class Errors, trigger "Défauts_Def_Canal02" bit 9
   19: 'Défaut Arret urgence', class Errors, trigger "Défauts_Def_Canal02" bit 10
   20: 'Défaut presence air', class Errors, trigger "Défauts_Def_Canal02" bit 11
   21: 'Défaut Robot 01', class Errors, trigger "Défauts_Def_Canal02" bit 12
   22: 'Défaut Robot 02', class Errors, trigger "Défauts_Def_Canal02" bit 13
   23: 'Défaut Robot 03', class Errors, trigger "Défauts_Def_Canal02" bit 14
   24: 'Défaut Robot 04', class Errors, trigger "Défauts_Def_Canal02" bit 15
   25: 'Défaut Robot 05', class Errors, trigger "Défauts_Def_Canal02" bit 0
   26: 'Défaut Vision', class Errors, trigger "Défauts_Def_Canal02" bit 1
   27: 'Défaut Axe Robot', class Errors, trigger "Défauts_Def_Canal02" bit 2
   28: '', class Errors, trigger "Défauts_Def_Canal02" bit 3
   29: '', class Errors, trigger "Défauts_Def_Canal02" bit 4
   30: '', class Errors, trigger "Défauts_Def_Canal02" bit 5
   31: '', class Errors, trigger "Défauts_Def_Canal02" bit 6
   32: '', class Errors, trigger "Défauts_Def_Canal02" bit 7
   33: 'Init_pas_possible_FANUC1_Pas_En_Auto', class Warnings, trigger "Défauts_Def_Canal03" bit 9
   34: 'Init_pas_possible_FANUC2_Pas_En_Auto', class Warnings, trigger "Défauts_Def_Canal03" bit 10
   35: 'Position finale non atteinte', class Warnings, trigger "Défauts_Def_Canal03" bit 11
   36: '', class Warnings, trigger "Défauts_Def_Canal03" bit 12

screen "Principale" 1280x800, template "Modèle_1"
   Button "Bouton_1" at 48,413 size 127x79; TextOff 'Depart Cycle'
      on Press: SetBit("Touche_Tch_DCY")
      on Release: ResetBit("Touche_Tch_DCY")
      Appearance <- "B_VOY_DCY"
      ObjectEnable <- "Bits_Globaux_x_En_auto"
   Button "Bouton_2" at 48,496 size 127x79; TextOff 'Arret Cycle'
      on Press: SetBit("Touche_Tch_FDCY")
      on Release: ResetBit("Touche_Tch_FDCY")
      Appearance <- "B_VOY_ACY"
   GraphicView "Vue de graphique_3" at 230,144 size 1023x553; Picture "Capture d’écran 2023-07-10 135110"
   TextField "Champ de texte_1" at 31,135 size 158x25; Text 'CDT DE MARCHE'
   Rectangle "Rectangle_8" at 29,158 size 24x24
      Appearance <- "I_En_Arret_Urgence"
   TextField "Champ de texte_2" at 55,159 size 143x25; Text 'Arret Urgence'
   Rectangle "Rectangle_9" at 29,186 size 24x24
      Appearance <- "Bits_Globaux_x_En_auto"
   TextField "Champ de texte_3" at 55,187 size 113x25; Text 'Mode Auto'
   Rectangle "Rectangle_10" at 29,214 size 24x24
      Appearance <- "I_En_Service"
   TextField "Champ de texte_4" at 61,215 size 103x25; Text 'En Service'
   Button "Bouton_3" at 1177,723 size 96x70; TextOff 'IN / OUT'
      on Release: ActivateScreen("Visu_ES-Cpu", 0)
   Button "Bouton_4" at 95,721 size 96x70; TextOff 'Alarmes'
      on Release: ActivateScreen("Alarmes", 0)
      Appearance <- "Bits_B_defaut_en_cours"
   GraphicView "Vue de graphique_5" at 19,728 size 60x60; Picture "Graphique_1"
      Visibility <- "Bits_B_defaut_en_cours"
   Button "Bouton_5" at 1070,723 size 96x70; TextOff 'PARAM'
      on Release: ActivateScreen("Parametrage", 0)
   Button "Bouton_6" at 963,723 size 96x70; TextOff 'MODE MANUEL'
      on Release: ActivateScreen("Mode_Manuel_B01_std_1", 0)
      ObjectEnable <- "Bits_Globaux_x_En_manu"
      Appearance <- "Bits_Globaux_x_En_manu"
   Button "Bouton_7" at 856,723 size 96x70; TextOff 'TP Robots'
      on Click: ActivateScreen("TP_Robots", 0)
      Appearance <- "B_Pret_TP_Robotique"
      on Release: InvertBit("Bits_B_TP_Robot")
   Button "Bouton_8" at 749,723 size 96x70; TextOff 'INIT.'
      on Press: SetBit("Touche_Tch_Init")
      on Release: ResetBit("Touche_Tch_Init")
      Appearance <- "VOY_Init"
      ObjectEnable <- "Bits_Globaux_x_Defaut_non_bloquant"
   Button "Bouton_10" at 535,723 size 96x70; TextOff 'AGVs'
      on Press: ActivateScreen("AGVs", 0)
   Button "Bouton_11" at 428,723 size 96x70; TextOff 'Text'
   Button "Bouton_12" at 321,723 size 96x70; TextOff 'Text'
   Button "Bouton_13" at 214,723 size 96x70; TextOff 'Acquit Defaut'
      on Press: SetBit("Touche_Tch_Acquit")
      on Release: ResetBit("Touche_Tch_Acquit")
   Circle "Cercle_1" at 473,447 size 28x28
      Appearance <- "Défauts_Defauts{0}"
      Visibility <- "Défauts_Defauts{0}"
   Circle "Cercle_2" at 358,447 size 28x28
      Appearance <- "Défauts_Defauts{1}"
      Visibility <- "Défauts_Defauts{1}"
   Circle "Cercle_3" at 266,512 size 28x28
      Appearance <- "Défauts_Defauts{2}"
      Visibility <- "Défauts_Defauts{2}"
   Circle "Cercle_4" at 412,565 size 28x28
      Visibility <- "Défauts_Defauts{12}"
      Appearance <- "Défauts_Defauts{12}"
   Circle "Cercle_5" at 629,564 size 28x28
      Appearance <- "Défauts_Defauts{13}"
      Visibility <- "Défauts_Defauts{13}"
   Circle "Cercle_6" at 760,504 size 28x28
      Visibility <- "Défauts_Defauts{14}"
      Appearance <- "Défauts_Defauts{14}"
   Circle "Cercle_7" at 615,447 size 28x28
      Appearance <- "Défauts_Defauts{15}"
      Visibility <- "Défauts_Defauts{15}"
   Circle "Cercle_8" at 775,565 size 28x28
      Visibility <- "Défauts_Defauts{3}"
      Appearance <- "Défauts_Defauts{3}"
   Circle "Cercle_9" at 760,437 size 28x28
      Appearance <- "Défauts_Defauts{4}"
      Visibility <- "Défauts_Defauts{4}"
   Circle "Cercle_10" at 262,447 size 28x28
      Visibility <- "Défauts_Defauts{5}"
      Appearance <- "Défauts_Defauts{5}"
   Circle "Cercle_11" at 262,571 size 28x28
      Appearance <- "Défauts_Defauts{6}"
      Visibility <- "Défauts_Defauts{6}"
   Circle "Cercle_12" at 963,392 size 28x28
      Visibility <- "Défauts_Defauts{7}"
      Appearance <- "Défauts_Defauts{7}"
   Circle "Cercle_13" at 1096,276 size 28x28
      Visibility <- "Défauts_Defauts{16}"
      Appearance <- "Défauts_Defauts{16}"
   Circle "Cercle_14" at 904,284 size 28x28
      Appearance <- "Défauts_Defauts{17}"
      Visibility <- "Défauts_Defauts{17}"
   Circle "Cercle_15" at 862,447 size 28x28
      Appearance <- "Défauts_Defauts{8}"
      Visibility <- "Défauts_Defauts{8}"
   Circle "Cercle_16" at 861,416 size 28x28
      Visibility <- "Défauts_Defauts{9}"
      Appearance <- "Défauts_Defauts{9}"
   Circle "Cercle_17" at 931,447 size 28x28
      Appearance <- "Défauts_Defauts{11}"
      Visibility <- "Défauts_Defauts{11}"
   Circle "Cercle_18" at 931,416 size 28x28
      Appearance <- "Défauts_Defauts{10}"
      Visibility <- "Défauts_Defauts{10}"
   Circle "Cercle_19" at 683,495 size 28x28
      Visibility <- "Défauts_Defauts{20}"
      Appearance <- "Défauts_Defauts{20}"
   Circle "Cercle_20" at 989,534 size 28x28
      Appearance <- "Défauts_Defauts{21}"
      Visibility <- "Défauts_Defauts{21}"
   Circle "Cercle_21" at 1050,284 size 28x28
      Appearance <- "Défauts_Defauts{22}"
      Visibility <- "Défauts_Defauts{22}"
   Circle "Cercle_22" at 1059,160 size 28x28
      Visibility <- "Défauts_Defauts{23}"
      Appearance <- "Défauts_Defauts{23}"
   Circle "Cercle_23" at 721,379 size 28x28
      Appearance <- "Défauts_Defauts{24}"
      Visibility <- "Défauts_Defauts{24}"
   Circle "Cercle_24" at 262,513 size 28x28
      Visibility <- "Défauts_Defauts{25}"
      Appearance <- "Défauts_Defauts{25}"
   Rectangle "Rectangle_1" at 825,454 size 20x20
      Appearance <- "I_det_Phot_01"
   Rectangle "Rectangle_2" at 975,454 size 20x20
      Appearance <- "I_det_Phot_02"
   Rectangle "Rectangle_3" at 1124,454 size 20x20
      Appearance <- "I_det_Phot_03"
   Rectangle "Rectangle_4" at 957,344 size 20x20
      Appearance <- "I_Det_Photo_7"
   Rectangle "Rectangle_12" at 862,344 size 20x20
      Appearance <- "I_Det_Photo_8"
   Rectangle "Rectangle_13" at 779,344 size 20x20
      Appearance <- "I_Det_Photo_9"
   Rectangle "Rectangle_14" at 1169,168 size 20x20
      Appearance <- "I_det_photo_03"
   Rectangle "Rectangle_15" at 1260,0 size 20x20
      Appearance <- "I_Det_Photo_9"
   Rectangle "Rectangle_16" at 1169,270 size 20x20
      Appearance <- "I_det_photo_02"
   Rectangle "Rectangle_17" at 1169,372 size 20x20
      Appearance <- "I_det_photo_01"
   Circle "Cercle_25" at 348,499 size 28x28
      Appearance <- "Défauts_Defauts{26}"
      Visibility <- "Défauts_Defauts{26}"
   Rectangle "Rectangle_18" at 29,242 size 24x24
      Appearance <- "I_Wieland_Porte 01 ouverte"
   TextField "Champ de texte_5" at 61,242 size 155x25; Text 'Porte Ouverte 1'
   Rectangle "Rectangle_19" at 29,270 size 24x24
      Appearance <- "I_Wieland_Porte 02 Ouverte"
   TextField "Champ de texte_6" at 61,270 size 155x25; Text 'Porte Ouverte 2'
   Rectangle "Rectangle_20" at 29,298 size 24x24
      Appearance <- "I_Wieland_Porte_non_Réarmée"
   TextField "Champ de texte_7" at 61,298 size 144x25; Text 'Porte Réarmée'
   TextField "Champ de texte_8" at 616,424 size 29x25; Text '01'
   TextField "Champ de texte_9" at 474,424 size 29x25; Text '02'
   TextField "Champ de texte_10" at 357,424 size 29x25; Text '03'
   TextField "Champ de texte_11" at 219,514 size 29x25; Text '04'
   TextField "Champ de texte_12" at 411,594 size 29x25; Text '05'
   TextField "Champ de texte_13" at 628,592 size 29x25; Text '06'
   TextField "Champ de texte_14" at 789,505 size 29x25; Text '07'
   Button "Bouton_14" at 4,5 size 124x122; TextOff 'Text'
      on Click: ActivateScreen("Page_demarrage", 0)
   TextField "Champ de texte_15" at 28,593 size 170x46; Text 'INITIALISATION EN COURS'
      Visibility <- "Bits_B_dmd_Init_robot"
      Appearance <- "Bits_B_dmd_Init_robot"
   TextField "Champ de texte_16" at 901,613 size 213x25; Text 'FANUC1 PAS EN AUTO'
      Appearance <- "FanucR1_In_auto"
      Visibility <- "FanucR1_In_auto"
   Button "Bouton_9" at 642,723 size 96x70; TextOff 'DEMO. HIPPO'
      on Release: InvertBit("Bits_B_Demo_Hyppo"); ResetBit("Bits_B_TP_Robot")
      ObjectEnable <- "Bits_Init_glob_OK"
      Appearance <- "Voyants_HMI_x_VOY_Demo_pret"
   TextField "Champ de texte_17" at 905,239 size 213x25; Text 'FANUC2 PAS EN AUTO'
      Appearance <- "FanucR2_In_Auto"
      Visibility <- "FanucR2_In_Auto"
   TextField "Champ de texte_18" at 902,592 size 205x25; Text 'FANUC1 Teach activé'
      Appearance <- "Fanuc1_Teach_active"
      Visibility <- "Fanuc1_Teach_active"
   TextField "Champ de texte_19" at 905,223 size 205x25; Text 'FANUC2 Teach activé'
      Appearance <- "Fanuc2_teach_active"
      Visibility <- "Fanuc2_teach_active"
   TextField "Champ de texte_20" at 231,187 size 234x25; Text 'Initialisation nécessaire'
      Appearance <- "Voyants_HMI_x_VOY_Init_requis_en_auto"
      Visibility <- "Voyants_HMI_x_VOY_Init_requis_en_auto"
   GraphicView "Graphic view_1" at 169,185 size 45x30; Picture "Graphic_7"
      Visibility <- "I_En_Automatique"
      Appearance <- "Bits_Globaux_x_En_auto"
   TextField "Champ de texte_21" at 231,227 size 213x25; Text 'FANUC1 PAS EN AUTO'
      Appearance <- "FanucR1_In_auto"
      Visibility <- "I_En_Automatique"
   TextField "Champ de texte_22" at 231,261 size 213x25; Text 'FANUC2 PAS EN AUTO'
      Appearance <- "FanucR2_In_Auto"
      Visibility <- "I_En_Automatique"
   TextField "Champ de texte_23" at 231,206 size 205x25; Text 'FANUC1 Teach activé'
      Appearance <- "Fanuc1_Teach_active"
      Visibility <- "I_En_Automatique"
   TextField "Champ de texte_24" at 231,245 size 205x25; Text 'FANUC2 Teach activé'
      Appearance <- "Fanuc2_teach_active"
      Visibility <- "I_En_Automatique"
   Button "Button_1" at 310,353 size 75x75; TextOff 'Text'; PictureOff "PrusaMK4-noBG"
      on Release: function_efd93a16("PopUp_Imp3d_1", 310, 50, -1, -1, 1)
   Button "Button_2" at 377,353 size 75x75; TextOff 'Text'; PictureOff "PrusaMK4-noBG"
      on Release: function_efd93a16("PopUp_Imp3d_2", 310, 50, -1, -1, 1)
   Button "Button_3" at 444,353 size 75x75; TextOff 'Text'; PictureOff "PrusaMK4-noBG"
      on Release: function_efd93a16("PopUp_Imp3d_3", 310, 50, -1, -1, 1)
   Button "Button_4" at 511,353 size 75x75; TextOff 'Text'; PictureOff "PrusaMK4-noBG"
      on Release: function_efd93a16("PopUp_Imp3d_4", 310, 50, -1, -1, 1)
   Rectangle "Rectangle_21" at 29,326 size 24x24
      Appearance <- "PW: Is power on"
   TextField "Champ de texte_25" at 61,327 size 115x25; Text 'UR4 Allumé'
   Rectangle "Rectangle_22" at 29,354 size 24x24
      Appearance <- "PW: Is power on"
   TextField "Champ de texte_26" at 61,355 size 115x25; Text 'UR5 Allumé'

screen "Page_demarrage" 1280x800
   GraphicView "Vue de graphique_1" at 243,0 size 800x800; Picture "unilasalle"
   Button "Bouton_1" at 6,5 size 1267x791; TextOff 'Text'
      on Click: ActivateScreen("Principale", 0)
   TextField "Champ de texte_1" at 820,743 size 443x29; Text 'Appuyer sur l'ecran pour demarrer ....'
   Switch "Switch_1" at 11,9 size 108x41; CaptionText 'Switch'; TextOff 'OFF'; TextOn 'ON'
      on Change: StopRuntime(0)

screen "Alarmes" 1280x800, template "Modèle_1"
   AlarmView "Vue des alarmes_1" at 14,132 size 1064x653
   Button "Bouton_3" at 1177,723 size 96x70; TextOff 'RETOUR'
      on Release: ActivateScreen("Principale", 0)

screen "Visu_ES-Cpu" 1280x800, template "Modèle_ES"
   GraphicView "Vue de graphique_1" at 24,140 size 272x158; Picture "Graphique_3"
   Rectangle "Rectangle_1" at 338,213 size 20x20
      Appearance <- "I_En_Service"
   TextField "Champ de texte_1" at 364,211 size 103x25; Text 'En Service'
   Rectangle "Rectangle_2" at 338,235 size 20x20
      Appearance <- "I_En_Arret_Urgence"
   TextField "Champ de texte_2" at 364,233 size 166x25; Text 'En Arret Urgence'
   Rectangle "Rectangle_3" at 338,257 size 20x20
      Appearance <- "I_En_Manuel"
   TextField "Champ de texte_3" at 364,255 size 102x25; Text 'En Manuel'
   Rectangle "Rectangle_4" at 338,279 size 20x20
      Appearance <- "I_En_Automatique"
   TextField "Champ de texte_4" at 364,277 size 156x25; Text 'En Automatique'
   Rectangle "Rectangle_5" at 338,301 size 20x20
      Appearance <- "I_porte_non_réarmée"
   TextField "Champ de texte_5" at 364,299 size 188x25; Text 'Porte Non Réarmée'
   Rectangle "Rectangle_6" at 338,323 size 20x20
      Appearance <- "I_porte_01_Op"
   TextField "Champ de texte_6" at 364,321 size 167x25; Text 'Porte 01 Ouverte'
   Rectangle "Rectangle_7" at 338,345 size 20x20
      Appearance <- "I_porte_02_Op"
   TextField "Champ de texte_7" at 364,343 size 167x25; Text 'Porte 02 Ouverte'
   Rectangle "Rectangle_8" at 338,367 size 20x20
      Appearance <- "I_libre_I07"
   TextField "Champ de texte_8" at 364,365 size 53x25; Text 'Libre'
   Rectangle "Rectangle_9" at 548,213 size 20x20
      Appearance <- "I_libre_I20"
   TextField "Champ de texte_9" at 574,211 size 53x25; Text 'Libre'
   Rectangle "Rectangle_10" at 548,235 size 20x20
      Appearance <- "I_libre_I21"
   TextField "Champ de texte_10" at 574,233 size 53x25; Text 'Libre'
   Rectangle "Rectangle_11" at 548,257 size 20x20
      Appearance <- "I_libre_I22"
   TextField "Champ de texte_11" at 574,255 size 53x25; Text 'Libre'
   Rectangle "Rectangle_12" at 548,279 size 20x20
      Appearance <- "I_libre_I23"
   TextField "Champ de texte_12" at 574,277 size 53x25; Text 'Libre'
   Rectangle "Rectangle_13" at 548,301 size 20x20
      Appearance <- "I_libre_I24"
   TextField "Champ de texte_13" at 574,299 size 53x25; Text 'Libre'
   Rectangle "Rectangle_14" at 548,323 size 20x20
      Appearance <- "I_libre_I25"
   TextField "Champ de texte_14" at 574,321 size 53x25; Text 'Libre'
   Rectangle "Rectangle_15" at 548,345 size 20x20
      Appearance <- "I_libre_I26"
   TextField "Champ de texte_15" at 574,343 size 53x25; Text 'Libre'
   Rectangle "Rectangle_16" at 548,367 size 20x20
      Appearance <- "I_libre_I27"
   TextField "Champ de texte_16" at 574,365 size 53x25; Text 'Libre'
   Rectangle "Rectangle_17" at 338,447 size 20x20
      Appearance <- "I_libre_I10"
   TextField "Champ de texte_17" at 364,445 size 53x25; Text 'Libre'
   Rectangle "Rectangle_18" at 338,469 size 20x20
      Appearance <- "I_Def_Thermique_CV01_hyppo"
   TextField "Champ de texte_18" at 364,467 size 159x25; Text 'Thermique CV01'
   Rectangle "Rectangle_19" at 338,491 size 20x20
      Appearance <- "I_Def_Thermique_CV02_hyppo"
   TextField "Champ de texte_19" at 364,489 size 159x25; Text 'Thermique CV02'
   Rectangle "Rectangle_20" at 338,513 size 20x20
      Appearance <- "I_Def_Thermique_CV03_hyppo"
   TextField "Champ de texte_20" at 364,511 size 159x25; Text 'Thermique CV03'
   Rectangle "Rectangle_21" at 338,535 size 20x20
      Appearance <- "I_Def_Thermique_CV04_hyppo"
   TextField "Champ de texte_21" at 364,533 size 159x25; Text 'Thermique CV04'
   Rectangle "Rectangle_22" at 338,557 size 20x20
      Appearance <- "I_libre_I15"
   TextField "Champ de texte_22" at 364,555 size 53x25; Text 'Libre'
   Rectangle "Rectangle_23" at 338,579 size 20x20
      Appearance <- "I_libre_I16"
   TextField "Champ de texte_23" at 364,577 size 53x25; Text 'Libre'
   Rectangle "Rectangle_24" at 338,601 size 20x20
      Appearance <- "I_libre_I17"
   TextField "Champ de texte_24" at 364,599 size 53x25; Text 'Libre'
   Rectangle "Rectangle_25" at 548,447 size 20x20
      Appearance <- "I_libre_I30"
   TextField "Champ de texte_25" at 574,445 size 53x25; Text 'Libre'
   Rectangle "Rectangle_26" at 548,469 size 20x20
      Appearance <- "I_libre_I31"
   TextField "Champ de texte_26" at 574,467 size 53x25; Text 'Libre'
   Rectangle "Rectangle_27" at 548,491 size 20x20
      Appearance <- "I_libre_I32"
   TextField "Champ de texte_27" at 574,489 size 53x25; Text 'Libre'
   Rectangle "Rectangle_28" at 548,513 size 20x20
      Appearance <- "I_libre_I33"
   TextField "Champ de texte_28" at 574,511 size 53x25; Text 'Libre'
   Rectangle "Rectangle_29" at 548,535 size 20x20
      Appearance <- "I_libre_I34"
   TextField "Champ de texte_29" at 574,533 size 53x25; Text 'Libre'
   Rectangle "Rectangle_30" at 548,557 size 20x20
      Appearance <- "I_libre_I35"
   TextField "Champ de texte_30" at 574,555 size 53x25; Text 'Libre'
   Rectangle "Rectangle_31" at 548,579 size 20x20
      Appearance <- "I_libre_I36"
   TextField "Champ de texte_31" at 574,577 size 53x25; Text 'Libre'
   Rectangle "Rectangle_32" at 548,601 size 20x20
      Appearance <- "I_libre_I37"
   TextField "Champ de texte_32" at 574,599 size 53x25; Text 'Libre'
   TextField "Champ de texte_33" at 319,142 size 459x25; Text 'ENTREES'
   TextField "Champ de texte_34" at 338,188 size 47x25; Text '%I0'
   TextField "Champ de texte_35" at 334,420 size 47x25; Text '%I1'
   TextField "Champ de texte_36" at 548,188 size 47x25; Text '%I2'
   TextField "Champ de texte_37" at 548,420 size 47x25; Text '%I3'
   Rectangle "Rectangle_36" at 813,213 size 20x20
      Appearance <- "Q_CL_verte"
   TextField "Champ de texte_38" at 839,211 size 138x25; Text 'Colonne Verte'
   Rectangle "Rectangle_37" at 813,235 size 20x20
      Appearance <- "Q_CL_Orange"
   TextField "Champ de texte_39" at 839,233 size 156x25; Text 'Colonne Orange'
   Rectangle "Rectangle_38" at 813,257 size 20x20
      Appearance <- "Q_CL_Rouge"
   TextField "Champ de texte_40" at 839,255 size 148x25; Text 'Colonne Rouge'
   Rectangle "Rectangle_39" at 813,279 size 20x20
      Appearance <- "Q_LibreQ03"
   TextField "Champ de texte_41" at 839,277 size 53x25; Text 'Libre'
   Rectangle "Rectangle_40" at 813,301 size 20x20
      Appearance <- "Q_LibreQ04"
   TextField "Champ de texte_42" at 839,299 size 53x25; Text 'Libre'
   Rectangle "Rectangle_41" at 813,323 size 20x20
      Appearance <- "Q_LibreQ05"
   TextField "Champ de texte_43" at 839,321 size 53x25; Text 'Libre'
   Rectangle "Rectangle_42" at 813,345 size 20x20
      Appearance <- "Q_LibreQ06"
   TextField "Champ de texte_44" at 839,343 size 53x25; Text 'Libre'
   Rectangle "Rectangle_43" at 813,367 size 20x20
      Appearance <- "Q_LibreQ07"
   TextField "Champ de texte_45" at 839,365 size 53x25; Text 'Libre'
   Rectangle "Rectangle_44" at 1023,213 size 20x20
      Appearance <- "Q_ON_CV_01_Hyppo"
   TextField "Champ de texte_46" at 1049,211 size 85x25; Text 'On CV01'
   Rectangle "Rectangle_45" at 1023,235 size 20x20
      Appearance <- "Q_ON_CV_02_Hyppo"
   TextField "Champ de texte_47" at 1049,233 size 85x25; Text 'On CV02'
   Rectangle "Rectangle_46" at 1023,257 size 20x20
      Appearance <- "Q_ON_CV_03_Hyppo"
   TextField "Champ de texte_48" at 1049,255 size 85x25; Text 'On CV03'
   Rectangle "Rectangle_47" at 1023,279 size 20x20
      Appearance <- "Q_ON_CV_04_Hyppo"
   TextField "Champ de texte_49" at 1049,277 size 84x25; Text 'On Cv04'
   Rectangle "Rectangle_48" at 1023,301 size 20x20
      Appearance <- "Q_LibreQ24"
   TextField "Champ de texte_50" at 1049,299 size 53x25; Text 'Libre'
   Rectangle "Rectangle_49" at 1023,323 size 20x20
      Appearance <- "Q_LibreQ25"
   TextField "Champ de texte_51" at 1049,321 size 53x25; Text 'Libre'
   Rectangle "Rectangle_50" at 1023,345 size 20x20
      Appearance <- "Q_LibreQ26"
   TextField "Champ de texte_52" at 1049,343 size 53x25; Text 'Libre'
   Rectangle "Rectangle_51" at 1023,367 size 20x20
      Appearance <- "Q_LibreQ27"
   TextField "Champ de texte_53" at 1049,365 size 53x25; Text 'Libre'
   Rectangle "Rectangle_52" at 813,447 size 20x20
      Appearance <- "Q_LibreQ10"
   TextField "Champ de texte_54" at 839,445 size 53x25; Text 'Libre'
   Rectangle "Rectangle_53" at 813,469 size 20x20
      Appearance <- "Q_LibreQ11"
   TextField "Champ de texte_55" at 839,467 size 53x25; Text 'Libre'
   Rectangle "Rectangle_54" at 813,491 size 20x20
      Appearance <- "Q_LibreQ12"
   TextField "Champ de texte_56" at 839,489 size 53x25; Text 'Libre'
   Rectangle "Rectangle_55" at 813,513 size 20x20
      Appearance <- "Q_LibreQ13"
   TextField "Champ de texte_57" at 839,511 size 53x25; Text 'Libre'
   Rectangle "Rectangle_56" at 813,535 size 20x20
      Appearance <- "Q_LibreQ14"
   TextField "Champ de texte_58" at 839,533 size 53x25; Text 'Libre'
   Rectangle "Rectangle_57" at 813,557 size 20x20
      Appearance <- "Q_LibreQ15"
   TextField "Champ de texte_59" at 839,555 size 53x25; Text 'Libre'
   Rectangle "Rectangle_58" at 813,579 size 20x20
      Appearance <- "Q_LibreQ16"
   TextField "Champ de texte_60" at 839,577 size 53x25; Text 'Libre'
   Rectangle "Rectangle_59" at 813,601 size 20x20
      Appearance <- "Q_LibreQ17"
   TextField "Champ de texte_61" at 839,599 size 53x25; Text 'Libre'
   Rectangle "Rectangle_60" at 1023,447 size 20x20
      Appearance <- "Q_LibreQ30"
   TextField "Champ de texte_62" at 1049,445 size 53x25; Text 'Libre'
   Rectangle "Rectangle_61" at 1023,469 size 20x20
      Appearance <- "Q_LibreQ31"
   TextField "Champ de texte_63" at 1049,467 size 53x25; Text 'Libre'
   Rectangle "Rectangle_62" at 1023,491 size 20x20
      Appearance <- "Q_LibreQ32"
   TextField "Champ de texte_64" at 1049,489 size 53x25; Text 'Libre'
   Rectangle "Rectangle_63" at 1023,513 size 20x20
      Appearance <- "Q_LibreQ33"
   TextField "Champ de texte_65" at 1049,511 size 53x25; Text 'Libre'
   Rectangle "Rectangle_64" at 1023,535 size 20x20
      Appearance <- "Q_LibreQ34"
   TextField "Champ de texte_66" at 1049,533 size 53x25; Text 'Libre'
   Rectangle "Rectangle_65" at 1023,557 size 20x20
      Appearance <- "Q_LibreQ35"
   TextField "Champ de texte_67" at 1049,555 size 53x25; Text 'Libre'
   Rectangle "Rectangle_66" at 1023,579 size 20x20
      Appearance <- "Q_LibreQ36"
   TextField "Champ de texte_68" at 1049,577 size 53x25; Text 'Libre'
   Rectangle "Rectangle_67" at 1023,601 size 20x20
      Appearance <- "Q_LibreQ37"
   TextField "Champ de texte_69" at 1049,599 size 53x25; Text 'Libre'
   TextField "Champ de texte_70" at 794,142 size 459x25; Text 'SORTIES'
   TextField "Champ de texte_71" at 813,188 size 52x25; Text '%Q0'
   TextField "Champ de texte_72" at 809,420 size 52x25; Text '%Q1'
   TextField "Champ de texte_73" at 1023,188 size 52x25; Text '%Q2'
   TextField "Champ de texte_74" at 1023,420 size 52x25; Text '%Q3'

Template "Modèle_1" 1280x800
   GraphicView "Vue de graphique_2" at 9,8 size 111x116; Picture "unilasalle"
   DateTimeField "Champ de date/heure_1" at 1133,29 size 131x34
   DateTimeField "Champ de date/heure_2" at 1152,65 size 99x34
   GraphicView "Vue de graphique_1" at 129,8 size 113x116; Picture "Ascodero"
   TextField "Champ de texte_5" at 634,54 size 173x28; Text 'Usine Ecole 4.0'
   Button "Bouton_14" at 4,5 size 124x122; TextOff 'Text'
      on Click: ActivateScreen("Page_demarrage", 0)

screen "Visu_ES_REP1_4" 1280x800, template "Modèle_ES"
   GraphicView "Vue de graphique_1" at 62,186 size 76x151; Picture "Graphique_4"
   TextField "Champ de texte_1" at 43,144 size 59x25; Text 'REP 1'
   GraphicView "Vue de graphique_2" at 62,454 size 76x151; Picture "Graphique_4"
   TextField "Champ de texte_18" at 43,412 size 59x25; Text 'REP 2'
   GraphicView "Vue de graphique_3" at 681,186 size 76x151; Picture "Graphique_4"
   TextField "Champ de texte_41" at 662,144 size 59x25; Text 'REP 3'
   Rectangle "Rectangle_41" at 808,244 size 20x20
      Appearance <- "AlwaysFALSE"
   TextField "Champ de texte_42" at 834,242 size 53x25; Text 'Libre'
   Rectangle "Rectangle_42" at 808,266 size 20x20
      Appearance <- "AlwaysFALSE"
   TextField "Champ de texte_43" at 834,264 size 53x25; Text 'Libre'
   Rectangle "Rectangle_43" at 808,288 size 20x20
      Appearance <- "AlwaysFALSE"
   TextField "Champ de texte_44" at 834,286 size 53x25; Text 'Libre'
   Rectangle "Rectangle_44" at 808,310 size 20x20
      Appearance <- "AlwaysFALSE"
   TextField "Champ de texte_45" at 834,308 size 53x25; Text 'Libre'
   Rectangle "Rectangle_45" at 808,332 size 20x20
      Appearance <- "AlwaysFALSE"
   TextField "Champ de texte_46" at 834,330 size 53x25; Text 'Libre'
   Rectangle "Rectangle_46" at 808,354 size 20x20
      Appearance <- "AlwaysFALSE"
   TextField "Champ de texte_47" at 834,352 size 53x25; Text 'Libre'
   Rectangle "Rectangle_47" at 808,376 size 20x20
      Appearance <- "AlwaysFALSE"
   TextField "Champ de texte_48" at 834,374 size 53x25; Text 'Libre'
   Rectangle "Rectangle_48" at 808,398 size 20x20
      Appearance <- "AlwaysFALSE"
   TextField "Champ de texte_49" at 834,396 size 53x25; Text 'Libre'
   Rectangle "Rectangle_49" at 1018,244 size 20x20
      Appearance <- "AlwaysFALSE"
   TextField "Champ de texte_50" at 1044,242 size 53x25; Text 'Libre'
   Rectangle "Rectangle_50" at 1018,266 size 20x20
      Appearance <- "AlwaysFALSE"
   TextField "Champ de texte_51" at 1044,264 size 53x25; Text 'Libre'
   Rectangle "Rectangle_51" at 1018,288 size 20x20
      Appearance <- "AlwaysFALSE"
   TextField "Champ de texte_52" at 1044,286 size 53x25; Text 'Libre'
   Rectangle "Rectangle_52" at 1018,310 size 20x20
      Appearance <- "AlwaysFALSE"
   TextField "Champ de texte_53" at 1044,308 size 53x25; Text 'Libre'
   Rectangle "Rectangle_53" at 1018,332 size 20x20
      Appearance <- "AlwaysFALSE"
   TextField "Champ de texte_54" at 1044,330 size 53x25; Text 'Libre'
   Rectangle "Rectangle_54" at 1018,354 size 20x20
      Appearance <- "AlwaysFALSE"
   TextField "Champ de texte_55" at 1044,352 size 53x25; Text 'Libre'
   Rectangle "Rectangle_55" at 1018,376 size 20x20
      Appearance <- "AlwaysFALSE"
   TextField "Champ de texte_56" at 1044,374 size 53x25; Text 'Libre'
   Rectangle "Rectangle_56" at 1018,398 size 20x20
      Appearance <- "AlwaysFALSE"
   TextField "Champ de texte_57" at 1044,396 size 53x25; Text 'Libre'
   TextField "Champ de texte_58" at 789,173 size 459x25; Text 'ENTREES'
   TextField "Champ de texte_59" at 808,219 size 47x25; Text '%I8'
   TextField "Champ de texte_60" at 1018,219 size 47x25; Text '%I9'
   GraphicView "Vue de graphique_4" at 681,454 size 76x151; Picture "Graphique_4"
   TextField "Champ de texte_61" at 662,412 size 59x25; Text 'REP 4'
   Rectangle "Rectangle_2" at 189,244 size 20x20
      Appearance <- "I_Pres_Elev_B01"
   TextField "Champ de texte_2" at 424,242 size 168x25; Text 'Presence pal B01'
   Rectangle "Rectangle_3" at 189,266 size 20x20
      Appearance <- "I_Elev_01_Haut"
   TextField "Champ de texte_3" at 209,242 size 178x25; Text 'Presence Elev B01'
   Rectangle "Rectangle_4" at 189,288 size 20x20
      Appearance <- "I_Pres_Elev_B02"
   TextField "Champ de texte_4" at 424,265 size 177x25; Text 'Elevateur Bas B01'
   Rectangle "Rectangle_5" at 189,310 size 20x20
      Appearance <- "I_Elev_02_Haut"
   TextField "Champ de texte_5" at 211,265 size 188x25; Text 'Elevateur Haut B01'
   Rectangle "Rectangle_6" at 189,332 size 20x20
      Appearance <- "I_Pres_Elev_B03"
   TextField "Champ de texte_6" at 424,287 size 168x25; Text 'Presence pal B02'
   Rectangle "Rectangle_7" at 189,354 size 20x20
      Appearance <- "I_Elev_03_Haut"
   TextField "Champ de texte_7" at 209,287 size 178x25; Text 'Presence Elev B02'
   Rectangle "Rectangle_8" at 189,376 size 20x20
      Appearance <- "I_Pres_Elev_B04"
   TextField "Champ de texte_8" at 424,308 size 177x25; Text 'Elevateur Bas B02'
   Rectangle "Rectangle_9" at 189,398 size 20x20
      Appearance <- "I_Elev_04_Haut"
   TextField "Champ de texte_9" at 209,308 size 188x25; Text 'Elevateur Haut B02'
   Rectangle "Rectangle_10" at 399,244 size 20x20
      Appearance <- "I_Pres_Pal_B01"
   TextField "Champ de texte_10" at 424,330 size 168x25; Text 'Presence pal B03'
   Rectangle "Rectangle_11" at 399,266 size 20x20
      Appearance <- "I_Elev_01_Bas"
   TextField "Champ de texte_11" at 211,330 size 178x25; Text 'Presence Elev B03'
   Rectangle "Rectangle_12" at 399,288 size 20x20
      Appearance <- "I_Pres_Pal_B02"
   TextField "Champ de texte_12" at 424,352 size 177x25; Text 'Elevateur Bas B03'
   Rectangle "Rectangle_13" at 399,310 size 20x20
      Appearance <- "I_Elev_02_Bas"
   TextField "Champ de texte_13" at 211,352 size 188x25; Text 'Elevateur Haut B03'
   Rectangle "Rectangle_14" at 399,332 size 20x20
      Appearance <- "I_Pres_Pal_B03"
   TextField "Champ de texte_14" at 424,374 size 168x25; Text 'Presence pal B04'
   Rectangle "Rectangle_15" at 399,354 size 20x20
      Appearance <- "I_Elev_03_Bas"
   TextField "Champ de texte_15" at 209,374 size 178x25; Text 'Presence Elev B04'
   Rectangle "Rectangle_16" at 399,376 size 20x20
      Appearance <- "I_Pres_Pal_B04"
   TextField "Champ de texte_16" at 424,395 size 177x25; Text 'Elevateur Bas B04'
   Rectangle "Rectangle_17" at 399,398 size 20x20
      Appearance <- "I_Elev_04_Bas"
   TextField "Champ de texte_17" at 211,395 size 188x25; Text 'Elevateur Haut B04'
   TextField "Champ de texte_34" at 170,173 size 459x25; Text 'ENTREES'
   TextField "Champ de texte_35" at 189,219 size 47x25; Text '%I4'
   TextField "Champ de texte_37" at 399,219 size 47x25; Text '%I5'
   Rectangle "Rectangle_20" at 189,512 size 20x20
      Appearance <- "I_Pres_Elev_B05"
   TextField "Champ de texte_19" at 421,510 size 168x25; Text 'Presence pal B05'
   Rectangle "Rectangle_21" at 189,534 size 20x20
      Appearance <- "I_Elev_05_Haut"
   TextField "Champ de texte_20" at 211,510 size 178x25; Text 'Presence Elev B05'
   Rectangle "Rectangle_22" at 189,556 size 20x20
      Appearance <- "I_Pres_Elev_B06"
   TextField "Champ de texte_21" at 421,532 size 177x25; Text 'Elevateur Bas B05'
   Rectangle "Rectangle_23" at 189,578 size 20x20
      Appearance <- "I_Elev_06_Haut"
   TextField "Champ de texte_22" at 211,532 size 188x25; Text 'Elevateur Haut B05'
   Rectangle "Rectangle_24" at 189,600 size 20x20
      Appearance <- "I_Pres_Elev_B07"
   TextField "Champ de texte_23" at 421,554 size 168x25; Text 'Presence pal B06'
   Rectangle "Rectangle_25" at 189,622 size 20x20
      Appearance <- "I_Elev_07_Haut"
   TextField "Champ de texte_24" at 211,554 size 178x25; Text 'Presence Elev B06'
   Rectangle "Rectangle_26" at 189,644 size 20x20
      Appearance <- "I_porte_vision_cl"
   TextField "Champ de texte_25" at 421,576 size 177x25; Text 'Elevateur Bas B06'
   Rectangle "Rectangle_27" at 189,666 size 20x20
      Appearance <- "AlwaysFALSE"
   TextField "Champ de texte_26" at 211,576 size 188x25; Text 'Elevateur Haut B06'
   Rectangle "Rectangle_28" at 399,512 size 20x20
      Appearance <- "I_Pres_Pal_B05"
   TextField "Champ de texte_27" at 421,598 size 168x25; Text 'Presence pal B07'
   Rectangle "Rectangle_29" at 399,534 size 20x20
      Appearance <- "I_Elev_05_Bas"
   TextField "Champ de texte_28" at 211,598 size 178x25; Text 'Presence Elev B07'
   Rectangle "Rectangle_30" at 399,556 size 20x20
      Appearance <- "I_Pres_Pal_B06"
   TextField "Champ de texte_29" at 421,620 size 177x25; Text 'Elevateur Bas B07'
   Rectangle "Rectangle_31" at 399,578 size 20x20
      Appearance <- "I_Elev_06_Bas"
   TextField "Champ de texte_30" at 211,620 size 188x25; Text 'Elevateur Haut B07'
   Rectangle "Rectangle_32" at 399,600 size 20x20
      Appearance <- "I_Pres_Pal_B07"
   TextField "Champ de texte_31" at 421,642 size 201x25; Text 'Porte Vision Ouverte'
   Rectangle "Rectangle_34" at 399,622 size 20x20
      Appearance <- "I_Elev_07_Bas"
   TextField "Champ de texte_32" at 211,642 size 192x25; Text 'Porte Vision fermée'
   Rectangle "Rectangle_36" at 399,644 size 20x20
      Appearance <- "I_porte_vision_op"
   TextField "Champ de texte_33" at 421,664 size 53x25; Text 'Libre'
   Rectangle "Rectangle_37" at 399,666 size 20x20
      Appearance <- "AlwaysFALSE"
   TextField "Champ de texte_36" at 211,664 size 53x25; Text 'Libre'
   TextField "Champ de texte_38" at 170,441 size 459x25; Text 'ENTREES'
   TextField "Champ de texte_39" at 189,487 size 47x25; Text '%I6'
   TextField "Champ de texte_40" at 399,487 size 47x25; Text '%I7'
   Rectangle "Rectangle_60" at 808,512 size 20x20
      Appearance <- "I_det_Phot_02"
   TextField "Champ de texte_62" at 1039,510 size 154x25; Text 'Det. Photo. N°1'
   Rectangle "Rectangle_61" at 808,534 size 20x20
      Appearance <- "I_verin_blocage_boite_sorti_01"
   TextField "Champ de texte_63" at 829,510 size 154x25; Text 'Det. Photo. N°2'
   Rectangle "Rectangle_62" at 808,556 size 20x20
      Appearance <- "I_verin_blocage_boite_sorti_02"
   TextField "Champ de texte_64" at 1039,532 size 154x25; Text 'Det. Photo. N°3'
   Rectangle "Rectangle_63" at 808,578 size 20x20
      Appearance <- "I_verin_blocage_boite_sorti_03"
   TextField "Champ de texte_65" at 829,532 size 182x25; Text 'Verin bloc 01 Sorti'
   Rectangle "Rectangle_64" at 808,600 size 20x20
      Appearance <- "I_verin_blocage_boite_sorti_04"
   TextField "Champ de texte_66" at 1039,554 size 199x25; Text 'Verin bloc 01 Rentré'
   Rectangle "Rectangle_65" at 808,622 size 20x20
      Appearance <- "AlwaysFALSE"
   TextField "Champ de texte_67" at 829,554 size 182x25; Text 'Verin bloc 02 Sorti'
   Rectangle "Rectangle_66" at 808,644 size 20x20
      Appearance <- "AlwaysFALSE"
   TextField "Champ de texte_68" at 1039,576 size 199x25; Text 'Verin bloc 02 Rentré'
   Rectangle "Rectangle_67" at 808,666 size 20x20
      Appearance <- "AlwaysFALSE"
   TextField "Champ de texte_69" at 829,575 size 182x25; Text 'Verin bloc 03 Sorti'
   Rectangle "Rectangle_68" at 1018,512 size 20x20
      Appearance <- "I_det_Phot_01"
   TextField "Champ de texte_70" at 1039,598 size 199x25; Text 'Verin bloc 03 Rentré'
   Rectangle "Rectangle_69" at 1018,534 size 20x20
      Appearance <- "I_det_Phot_03"
   TextField "Champ de texte_71" at 829,598 size 182x25; Text 'Verin bloc 04 Sorti'
   Rectangle "Rectangle_70" at 1018,556 size 20x20
      Appearance <- "I_verin_blocage_boite_rentré_01"
   TextField "Champ de texte_72" at 1039,620 size 199x25; Text 'Verin bloc 04 Rentré'
   Rectangle "Rectangle_71" at 1018,578 size 20x20
      Appearance <- "I_verin_blocage_boite_rentré_02"
   TextField "Champ de texte_73" at 829,621 size 53x25; Text 'Libre'
   TextField "Champ de texte_74" at 1039,642 size 53x25; Text 'Libre'
   Rectangle "Rectangle_73" at 1018,622 size 20x20
      Appearance <- "I_verin_blocage_boite_rentré_04"
   TextField "Champ de texte_75" at 829,643 size 53x25; Text 'Libre'
   Rectangle "Rectangle_74" at 1018,644 size 20x20
      Appearance <- "AlwaysFALSE"
   TextField "Champ de texte_76" at 1039,664 size 53x25; Text 'Libre'
   Rectangle "Rectangle_75" at 1018,666 size 20x20
      Appearance <- "AlwaysFALSE"
   TextField "Champ de texte_77" at 829,665 size 53x25; Text 'Libre'
   TextField "Champ de texte_78" at 789,441 size 459x25; Text 'ENTREES'
   TextField "Champ de texte_79" at 808,487 size 59x25; Text '%I10'
   TextField "Champ de texte_80" at 1018,487 size 59x25; Text '%I11'

Template "Modèle_ES" 1280x800
   Button "Bouton_5" at 861,723 size 96x70; TextOff 'Text'
   Button "Bouton_6" at 754,723 size 96x70; TextOff 'FANUC'
      on Click: ActivateScreen("Visu_ES-Fanuc", 0)
   Button "Bouton_7" at 647,723 size 96x70; TextOff 'VARIAT. G120C'
      on Release: ActivateScreen("Visu_ES_Variateur_C1", 0)
   Button "Bouton_8" at 540,723 size 96x70; TextOff 'WIELAND SECU.'
      on Release: ActivateScreen("Visu_ES_Wieland", 0)
   Button "Bouton_9" at 433,723 size 96x70; TextOff 'DISTRIB. ILOT02'
      on Release: ActivateScreen("Visu_ES_Ilot02", 0)
   Button "Bouton_10" at 326,723 size 96x70; TextOff 'DISTRIB. ILOT 01'
      on Release: ActivateScreen("Visu_ES_Ilot01", 0)
   Button "Bouton_11" at 219,723 size 96x70; TextOff 'REPART. RP5..6'
      on Release: ActivateScreen("Visu_ES_rep5_6", 0)
   Button "Bouton_12" at 112,723 size 96x70; TextOff 'REPART. RP1..4'
      on Release: ActivateScreen("Visu_ES_REP1_4", 0)
   Button "Bouton_13" at 5,723 size 96x70; TextOff 'CPU'
      on Release: ActivateScreen("Visu_ES-Cpu", 0)
   DateTimeField "Champ de date/heure_1" at 1133,29 size 131x34
   DateTimeField "Champ de date/heure_2" at 1152,65 size 99x34
   GraphicView "Vue de graphique_1" at 129,8 size 113x116; Picture "Ascodero"
   TextField "Champ de texte_5" at 600,51 size 172x28; Text 'Usine Ecole 4.0'
   GraphicView "Vue de graphique_2" at 9,8 size 111x116; Picture "unilasalle"
   Button "Bouton_3" at 1177,723 size 96x70; TextOff 'RETOUR'
      on Release: ActivateScreen("Principale", 0)
   Button "Bouton_1" at 1074,723 size 96x70; TextOff 'Text'
   Button "Bouton_2" at 967,723 size 96x70; TextOff 'Text'
   Button "Bouton_14" at 4,5 size 124x122; TextOff 'Text'
      on Click: ActivateScreen("Page_demarrage", 0)

